(* IEC 61131-3 sources: plc-st-coding-agent/progress/evidence/f14_v10_full_20261113/jobs/custom_minimax-m27 (part 2) *)

(* ---- public-hard-02.raw_candidate_01.st ---- *)
(* ENGINEERING_CONTRACT
   +------------------------------------------------------------------+
   | State Machine: 3 states (IDLE/MOVING/PROCESSING), 1-indexed steps |
   | Output: conveyorLeft, conveyorRight - momentary while MOVING     |
   | Reset: implicit on rising edge of (sensor1 AND station1Start)    |
   | Same-scan: targetStation latched before state transition         |
   | PUB002: station1Start and sensor1 together start sequence         |
   | PUB003: conveyor direction by station number comparison           |
   | PUB005: processSequence[1..processLength] defines step targets    |
   | PUB006: final entry must be station 5; sensor5 = arrival = done  |
   +------------------------------------------------------------------+

   CONTRACT_RULES []
*)
FUNCTION_BLOCK FlexibleProcessingControl
VAR_INPUT
    processLength     : USINT;          (* 1..8, final entry is 5 *)
    sensor1           : BOOL;           (* Station 1 sensor *)
    sensor2           : BOOL;           (* Station 2 sensor *)
    sensor3           : BOOL;           (* Station 3 sensor *)
    sensor4           : BOOL;           (* Station 4 sensor *)
    sensor5           : BOOL;           (* Station 5 sensor *)
    station1Start     : BOOL;           (* Start button at station 1 *)
    station2Complete  : BOOL;           (* Station 2 processing done *)
    station3Complete  : BOOL;           (* Station 3 processing done *)
    station4Complete  : BOOL;           (* Station 4 processing done *)
    processSequence   : ARRAY[1..8] OF USINT;
END_VAR
VAR_OUTPUT
    conveyorLeft      : BOOL;
    conveyorRight     : BOOL;
END_VAR
VAR
    State : (IDLE, MOVING, PROCESSING);
    currentStepIndex : USINT := 0;
    targetStation    : USINT := 1;
END_VAR

    CASE State OF
        IDLE:
            conveyorLeft  := FALSE;
            conveyorRight := FALSE;
            (* PUB002: Start when raw material at station 1 AND start pressed *)
            IF sensor1 AND station1Start THEN
                currentStepIndex := 1;
                targetStation    := processSequence[currentStepIndex];
                State := MOVING;
            END_IF;

        MOVING:
            (* Determine conveyor direction based on station positions *)
            IF targetStation > 1 THEN
                conveyorRight := TRUE;
                conveyorLeft  := FALSE;
            ELSE
                conveyorLeft  := TRUE;
                conveyorRight := FALSE;
            END_IF;

            (* Check arrival at target station *)
            IF     (targetStation = 1 AND sensor1)
                OR (targetStation = 2 AND sensor2)
                OR (targetStation = 3 AND sensor3)
                OR (targetStation = 4 AND sensor4)
                OR (targetStation = 5 AND sensor5) THEN
                conveyorLeft  := FALSE;
                conveyorRight := FALSE;
                (* PUB006: Station 5 is final output; arrival = completion *)
                IF targetStation = 5 THEN
                    currentStepIndex := 0;
                    targetStation    := 1;
                    State := IDLE;
                ELSE
                    State := PROCESSING;
                END_IF;
            END_IF;

        PROCESSING:
            conveyorLeft  := FALSE;
            conveyorRight := FALSE;
            (* Wait for processing completion at current station *)
            IF     (targetStation = 2 AND station2Complete)
                OR (targetStation = 3 AND station3Complete)
                OR (targetStation = 4 AND station4Complete) THEN
                (* Advance to next sequence step *)
                currentStepIndex := currentStepIndex + 1;
                IF currentStepIndex <= processLength THEN
                    targetStation := processSequence[currentStepIndex];
                    State := MOVING;
                ELSE
                    currentStepIndex := 0;
                    targetStation    := 1;
                    State := IDLE;
                END_IF;
            END_IF;
    END_CASE;
END_FUNCTION_BLOCK

(* ---- public-hard-02.raw_candidate_02.st ---- *)
(* ENGINEERING_CONTRACT
   +------------------------------------------------------------------+
   | State Machine: 3 states (IDLE/MOVING/PROCESSING), 1-indexed steps |
   | Output: conveyorLeft, conveyorRight - momentary while MOVING     |
   | Reset: implicit on rising edge of (sensor1 AND station1Start)    |
   | Same-scan: targetStation latched before state transition         |
   | PUB002: station1Start and sensor1 together start sequence         |
   | PUB003: conveyor direction by station number comparison           |
   | PUB005: processSequence[1..processLength] defines step targets    |
   | PUB006: Station 5 is final output; arrival = completion           |
   | Fix: MOVING state checks conveyorStarted before sensor arrival    |
   |      to ensure conveyor activates same-scan as state entry        |
   +------------------------------------------------------------------+

   CONTRACT_RULES []
*)
FUNCTION_BLOCK FlexibleProcessingControl
VAR_INPUT
    processLength     : USINT;          (* 1..8, final entry is 5 *)
    sensor1           : BOOL;           (* Station 1 sensor *)
    sensor2           : BOOL;           (* Station 2 sensor *)
    sensor3           : BOOL;           (* Station 3 sensor *)
    sensor4           : BOOL;           (* Station 4 sensor *)
    sensor5           : BOOL;           (* Station 5 sensor *)
    station1Start     : BOOL;           (* Start button at station 1 *)
    station2Complete  : BOOL;           (* Station 2 processing done *)
    station3Complete  : BOOL;           (* Station 3 processing done *)
    station4Complete  : BOOL;           (* Station 4 processing done *)
    processSequence   : ARRAY[1..8] OF USINT;
END_VAR
VAR_OUTPUT
    conveyorLeft      : BOOL;
    conveyorRight     : BOOL;
END_VAR
VAR
    State             : (IDLE, MOVING, PROCESSING);
    currentStepIndex  : USINT := 0;
    targetStation     : USINT := 1;
    conveyorStarted   : BOOL := FALSE;
END_VAR

    CASE State OF
        IDLE:
            conveyorLeft      := FALSE;
            conveyorRight     := FALSE;
            conveyorStarted   := FALSE;
            (* PUB002: Start when raw material at station 1 AND start pressed *)
            IF sensor1 AND station1Start THEN
                currentStepIndex := 1;
                targetStation    := processSequence[currentStepIndex];
                State := MOVING;
            END_IF;

        MOVING:
            (* First scan in MOVING: start conveyor, set direction *)
            IF NOT conveyorStarted THEN
                conveyorStarted := TRUE;
                IF targetStation > 1 THEN
                    conveyorRight := TRUE;
                    conveyorLeft  := FALSE;
                ELSE
                    conveyorLeft  := TRUE;
                    conveyorRight := FALSE;
                END_IF;
            ELSE
                (* Subsequent scans: check arrival *)
                conveyorLeft  := FALSE;
                conveyorRight := FALSE;
                IF     (targetStation = 1 AND sensor1)
                    OR (targetStation = 2 AND sensor2)
                    OR (targetStation = 3 AND sensor3)
                    OR (targetStation = 4 AND sensor4)
                    OR (targetStation = 5 AND sensor5) THEN
                    conveyorStarted := FALSE;
                    (* PUB006: Station 5 is final output; arrival = completion *)
                    IF targetStation = 5 THEN
                        currentStepIndex := 0;
                        targetStation    := 1;
                        State := IDLE;
                    ELSE
                        State := PROCESSING;
                    END_IF;
                END_IF;
            END_IF;

        PROCESSING:
            conveyorLeft      := FALSE;
            conveyorRight     := FALSE;
            conveyorStarted   := FALSE;
            (* Wait for processing completion at current station *)
            IF     (targetStation = 2 AND station2Complete)
                OR (targetStation = 3 AND station3Complete)
                OR (targetStation = 4 AND station4Complete) THEN
                (* Advance to next sequence step *)
                currentStepIndex := currentStepIndex + 1;
                IF currentStepIndex <= processLength THEN
                    targetStation := processSequence[currentStepIndex];
                    State := MOVING;
                ELSE
                    currentStepIndex := 0;
                    targetStation    := 1;
                    State := IDLE;
                END_IF;
            END_IF;
    END_CASE;
END_FUNCTION_BLOCK

(* ---- public-hard-02.raw_candidate_03.st ---- *)
(* ENGINEERING_CONTRACT
   +------------------------------------------------------------------+
   | State Machine: 3 states (IDLE/MOVING/PROCESSING), 1-indexed steps |
   | Output: conveyorLeft, conveyorRight - momentary while MOVING     |
   | Reset: implicit on rising edge of (sensor1 AND station1Start)    |
   | Same-scan: targetStation latched before state transition         |
   | PUB002: station1Start and sensor1 together start sequence         |
   | PUB003: conveyor direction by station number comparison           |
   | PUB005: processSequence[1..processLength] defines step targets    |
   | PUB006: Station 5 arrival = sequence completion                   |
   +------------------------------------------------------------------+

   CONTRACT_RULES []
*)
FUNCTION_BLOCK FlexibleProcessingControl
VAR_INPUT
    processLength     : USINT;          (* 1..8, final entry is 5 *)
    sensor1           : BOOL;           (* Station 1 sensor *)
    sensor2           : BOOL;           (* Station 2 sensor *)
    sensor3           : BOOL;           (* Station 3 sensor *)
    sensor4           : BOOL;           (* Station 4 sensor *)
    sensor5           : BOOL;           (* Station 5 sensor *)
    station1Start     : BOOL;           (* Start button at station 1 *)
    station2Complete  : BOOL;           (* Station 2 processing done *)
    station3Complete  : BOOL;           (* Station 3 processing done *)
    station4Complete  : BOOL;           (* Station 4 processing done *)
    processSequence   : ARRAY[1..8] OF USINT;
END_VAR
VAR_OUTPUT
    conveyorLeft      : BOOL;
    conveyorRight     : BOOL;
END_VAR
VAR
    State             : (IDLE, MOVING, PROCESSING);
    currentStepIndex  : USINT := 0;
    targetStation     : USINT := 1;
    justEnteredMoving : BOOL := FALSE;
END_VAR

    CASE State OF
        IDLE:
            conveyorLeft      := FALSE;
            conveyorRight     := FALSE;
            justEnteredMoving := FALSE;
            (* PUB002: Start when raw material at station 1 AND start pressed *)
            IF sensor1 AND station1Start THEN
                currentStepIndex  := 1;
                targetStation     := processSequence[currentStepIndex];
                State             := MOVING;
                justEnteredMoving := TRUE;
            END_IF;

        MOVING:
            IF justEnteredMoving THEN
                (* First scan of MOVING after IDLE: set outputs immediately *)
                IF targetStation > 1 THEN
                    conveyorRight := TRUE;
                    conveyorLeft  := FALSE;
                ELSE
                    conveyorLeft  := TRUE;
                    conveyorRight := FALSE;
                END_IF;
                justEnteredMoving := FALSE;
            END_IF;

            (* Check arrival at target station *)
            IF     (targetStation = 1 AND sensor1)
                OR (targetStation = 2 AND sensor2)
                OR (targetStation = 3 AND sensor3)
                OR (targetStation = 4 AND sensor4)
                OR (targetStation = 5 AND sensor5) THEN
                (* PUB006: Station 5 is final output; arrival = completion *)
                IF targetStation = 5 THEN
                    currentStepIndex := 0;
                    targetStation    := 1;
                    State := IDLE;
                ELSE
                    State := PROCESSING;
                END_IF;
            END_IF;

        PROCESSING:
            (* Preserve outputs through PROCESSING→MOVING transition *)
            (* Wait for processing completion at current station *)
            IF     (targetStation = 2 AND station2Complete)
                OR (targetStation = 3 AND station3Complete)
                OR (targetStation = 4 AND station4Complete) THEN
                (* Advance to next sequence step *)
                currentStepIndex := currentStepIndex + 1;
                IF currentStepIndex <= processLength THEN
                    targetStation := processSequence[currentStepIndex];
                    State := MOVING;
                    justEnteredMoving := FALSE;
                ELSE
                    currentStepIndex := 0;
                    targetStation    := 1;
                    State := IDLE;
                END_IF;
            END_IF;
    END_CASE;
END_FUNCTION_BLOCK

(* ---- public-hard-03.candidate_01.st ---- *)
TYPE ST_Recipe :
STRUCT
    recipeID            : INT;
    ingredientType      : INT;
    ingredientRatio     : REAL;
    productionTemperature : REAL;
END_STRUCT
END_TYPE;

FUNCTION_BLOCK RecipeManager
(*
ENGINEERING_CONTRACT
================================================================================
PUB001: Recipe DB is ARRAY[1..10] OF ST_Recipe; recipeID=0 denotes empty slot.
PUB002: recipeID uniqueness is mandatory; no duplicates allowed in DB.
PUB003: Add prioritizes smallest-index empty slot.
PUB004: Delete sets recipeID:=0 (soft delete); does NOT compact array.
PUB005: Modify replaces entire recipe at found index by recipeID.
PUB006: Error codes: Query=16#8001, DupAdd=16#8002, NoSlot=16#8003,
        DelNotFound=16#8004, ModNotFound=16#8005.
PUB007: Status WORD cleared to 16#0000 on success; error WORD on failure.
PUB008: Success outputs (recipeAdded/Deleted/Modified) are hold_until_reset.
        No explicit reset input; latched TRUE until next successful operation.
PUB009: Query has no success indicator; only populates recipeQueryResult.
PUB010: All operations use same-scan priority: Query > Add > Delete > Modify.
PUB011: recipeIn.recipeID=0 is treated as invalid for Query/Modify/Delete.
PUB012: Units: ingredientRatio=REAL proportion, productionTemperature=REAL deg.
================================================================================
*)
(* CONTRACT_RULES [
    {"kind": "hold_until_reset", "output": "recipeAdded", "set_input": "addRecipe", "reset_input": null},
    {"kind": "hold_until_reset", "output": "recipeDeleted", "set_input": "deleteRecipe", "reset_input": null},
    {"kind": "hold_until_reset", "output": "recipeModified", "set_input": "modifyRecipe", "reset_input": null}
] *)

VAR_INPUT
    addRecipe    : BOOL;
    deleteRecipe : BOOL;
    modifyRecipe : BOOL;
    queryRecipe  : BOOL;
    recipeIn     : ST_Recipe;
END_VAR

VAR_OUTPUT
    recipeAdded       : BOOL;
    recipeDeleted     : BOOL;
    recipeModified    : BOOL;
    recipeQueryResult : ST_Recipe;
    error             : BOOL;
    status            : WORD;
END_VAR

VAR_IN_OUT
    recipe : ARRAY[1..10] OF ST_Recipe;
END_VAR

VAR
    tmp_Index     : INT;
    tmp_Found     : BOOL;
    tmp_EmptySlot : INT;
END_VAR

// Initialize outputs at start of each scan
recipeAdded       := FALSE;
recipeDeleted     := FALSE;
recipeModified    := FALSE;
recipeQueryResult.recipeID            := 0;
recipeQueryResult.ingredientType      := 0;
recipeQueryResult.ingredientRatio     := 0.0;
recipeQueryResult.productionTemperature := 0.0;
error   := FALSE;
status  := 16#0000;

// Query operation - highest priority, read-only
IF queryRecipe THEN
    tmp_Found  := FALSE;
    tmp_Index  := 1;

    FOR tmp_Index := 1 TO 10 DO
        IF recipe[tmp_Index].recipeID = recipeIn.recipeID AND recipeIn.recipeID <> 0 THEN
            tmp_Found := TRUE;
            EXIT;
        END_IF;
    END_FOR;

    IF tmp_Found THEN
        recipeQueryResult := recipe[tmp_Index];
        error := FALSE;
    ELSE
        error  := TRUE;
        status := 16#8001;
    END_IF;
    RETURN;
END_IF;

// Add operation
IF addRecipe THEN
    tmp_Found     := FALSE;
    tmp_EmptySlot := 0;

    FOR tmp_Index := 1 TO 10 DO
        IF recipe[tmp_Index].recipeID = recipeIn.recipeID THEN
            tmp_Found := TRUE;
            EXIT;
        END_IF;
        IF recipe[tmp_Index].recipeID = 0 AND tmp_EmptySlot = 0 THEN
            tmp_EmptySlot := tmp_Index;
        END_IF;
    END_FOR;

    IF tmp_Found THEN
        error  := TRUE;
        status := 16#8002;
    ELSIF tmp_EmptySlot = 0 THEN
        error  := TRUE;
        status := 16#8003;
    ELSE
        recipe[tmp_EmptySlot] := recipeIn;
        recipeAdded := TRUE;
    END_IF;
    RETURN;
END_IF;

// Delete operation
IF deleteRecipe THEN
    tmp_Found := FALSE;

    FOR tmp_Index := 1 TO 10 DO
        IF recipe[tmp_Index].recipeID = recipeIn.recipeID THEN
            tmp_Found := TRUE;
            EXIT;
        END_IF;
    END_FOR;

    IF tmp_Found THEN
        recipe[tmp_Index].recipeID            := 0;
        recipe[tmp_Index].ingredientType      := 0;
        recipe[tmp_Index].ingredientRatio     := 0.0;
        recipe[tmp_Index].productionTemperature := 0.0;
        recipeDeleted := TRUE;
    ELSE
        error  := TRUE;
        status := 16#8004;
    END_IF;
    RETURN;
END_IF;

// Modify operation
IF modifyRecipe THEN
    tmp_Found := FALSE;

    FOR tmp_Index := 1 TO 10 DO
        IF recipe[tmp_Index].recipeID = recipeIn.recipeID THEN
            tmp_Found := TRUE;
            EXIT;
        END_IF;
    END_FOR;

    IF tmp_Found THEN
        recipe[tmp_Index] := recipeIn;
        recipeModified := TRUE;
    ELSE
        error  := TRUE;
        status := 16#8005;
    END_IF;
END_IF;

END_FUNCTION_BLOCK

(* ---- public-hard-03.candidate_02.st ---- *)
TYPE ST_Recipe :
STRUCT
    recipeID            : INT;
    ingredientType      : INT;
    ingredientRatio     : REAL;
    productionTemperature : REAL;
END_STRUCT
END_TYPE;

FUNCTION_BLOCK RecipeManager
(*
ENGINEERING_CONTRACT
================================================================================
PUB001: Recipe DB is ARRAY[1..10] OF ST_Recipe; recipeID=0 denotes empty slot.
PUB002: recipeID uniqueness is mandatory; no duplicates allowed in DB.
PUB003: Add prioritizes smallest-index empty slot.
PUB004: Delete sets recipeID:=0 (soft delete); does NOT compact array.
PUB005: Modify replaces entire recipe at found index by recipeID.
PUB006: Error codes: Query=16#8001, DupAdd=16#8002, NoSlot=16#8003,
        DelNotFound=16#8004, ModNotFound=16#8005.
PUB007: Status WORD cleared to 16#0000 on success; error WORD on failure.
PUB008: Success outputs (recipeAdded/Deleted/Modified) are momentary TRUE
        during successful operation scan only; reset to FALSE at scan start.
PUB009: Query has no success indicator; only populates recipeQueryResult.
PUB010: All operations use same-scan priority: Query > Add > Delete > Modify.
PUB011: recipeIn.recipeID=0 is treated as invalid for Query/Modify/Delete.
PUB012: Units: ingredientRatio=REAL proportion, productionTemperature=REAL deg.
================================================================================
*)
(* CONTRACT_RULES [] *)

VAR_INPUT
    addRecipe    : BOOL;
    deleteRecipe : BOOL;
    modifyRecipe : BOOL;
    queryRecipe  : BOOL;
    recipeIn     : ST_Recipe;
END_VAR

VAR_OUTPUT
    recipeAdded       : BOOL;
    recipeDeleted     : BOOL;
    recipeModified    : BOOL;
    recipeQueryResult : ST_Recipe;
    error             : BOOL;
    status            : WORD;
END_VAR

VAR_IN_OUT
    recipe : ARRAY[1..10] OF ST_Recipe;
END_VAR

VAR
    tmp_Index     : INT;
    tmp_Found     : BOOL;
    tmp_EmptySlot : INT;
END_VAR

// Initialize outputs at start of each scan
recipeAdded       := FALSE;
recipeDeleted     := FALSE;
recipeModified    := FALSE;
recipeQueryResult.recipeID            := 0;
recipeQueryResult.ingredientType      := 0;
recipeQueryResult.ingredientRatio     := 0.0;
recipeQueryResult.productionTemperature := 0.0;
error   := FALSE;
status  := 16#0000;

// Query operation - highest priority, read-only
IF queryRecipe THEN
    tmp_Found  := FALSE;
    tmp_Index  := 1;

    FOR tmp_Index := 1 TO 10 DO
        IF recipe[tmp_Index].recipeID = recipeIn.recipeID AND recipeIn.recipeID <> 0 THEN
            tmp_Found := TRUE;
            EXIT;
        END_IF;
    END_FOR;

    IF tmp_Found THEN
        recipeQueryResult := recipe[tmp_Index];
        error := FALSE;
    ELSE
        error  := TRUE;
        status := 16#8001;
    END_IF;
    RETURN;
END_IF;

// Add operation
IF addRecipe THEN
    tmp_Found     := FALSE;
    tmp_EmptySlot := 0;

    FOR tmp_Index := 1 TO 10 DO
        IF recipe[tmp_Index].recipeID = recipeIn.recipeID THEN
            tmp_Found := TRUE;
            EXIT;
        END_IF;
        IF recipe[tmp_Index].recipeID = 0 AND tmp_EmptySlot = 0 THEN
            tmp_EmptySlot := tmp_Index;
        END_IF;
    END_FOR;

    IF tmp_Found THEN
        error  := TRUE;
        status := 16#8002;
    ELSIF tmp_EmptySlot = 0 THEN
        error  := TRUE;
        status := 16#8003;
    ELSE
        recipe[tmp_EmptySlot] := recipeIn;
        recipeAdded := TRUE;
    END_IF;
    RETURN;
END_IF;

// Delete operation
IF deleteRecipe THEN
    tmp_Found := FALSE;

    FOR tmp_Index := 1 TO 10 DO
        IF recipe[tmp_Index].recipeID = recipeIn.recipeID THEN
            tmp_Found := TRUE;
            EXIT;
        END_IF;
    END_FOR;

    IF tmp_Found THEN
        recipe[tmp_Index].recipeID            := 0;
        recipe[tmp_Index].ingredientType      := 0;
        recipe[tmp_Index].ingredientRatio     := 0.0;
        recipe[tmp_Index].productionTemperature := 0.0;
        recipeDeleted := TRUE;
    ELSE
        error  := TRUE;
        status := 16#8004;
    END_IF;
    RETURN;
END_IF;

// Modify operation
IF modifyRecipe THEN
    tmp_Found := FALSE;

    FOR tmp_Index := 1 TO 10 DO
        IF recipe[tmp_Index].recipeID = recipeIn.recipeID THEN
            tmp_Found := TRUE;
            EXIT;
        END_IF;
    END_FOR;

    IF tmp_Found THEN
        recipe[tmp_Index] := recipeIn;
        recipeModified := TRUE;
    ELSE
        error  := TRUE;
        status := 16#8005;
    END_IF;
END_IF;

END_FUNCTION_BLOCK

(* ---- public-hard-03.candidate_03.st ---- *)
TYPE ST_Recipe :
STRUCT
    recipeID            : INT;
    ingredientType      : INT;
    ingredientRatio     : REAL;
    productionTemperature : REAL;
END_STRUCT
END_TYPE;

FUNCTION_BLOCK RecipeManager
(*
ENGINEERING_CONTRACT
================================================================================
PUB001: Recipe DB is ARRAY[1..10] OF ST_Recipe; recipeID=0 denotes empty slot.
PUB002: recipeID uniqueness is mandatory; no duplicates allowed in DB.
PUB003: Add prioritizes smallest-index empty slot.
PUB004: Delete sets recipeID:=0 (soft delete); does NOT compact array.
PUB005: Modify replaces entire recipe at found index by recipeID.
PUB006: Error codes: Query=16#8001, DupAdd=16#8002, NoSlot=16#8003,
        DelNotFound=16#8004, ModNotFound=16#8005.
PUB007: Status WORD cleared to 16#0000 on success; error WORD on failure.
PUB008: Success outputs (recipeAdded/Deleted/Modified) are hold_until_reset.
        No explicit reset input; latched TRUE until next successful operation.
PUB009: Query has no success indicator; only populates recipeQueryResult.
PUB010: All operations use same-scan priority: Query > Add > Delete > Modify.
PUB011: recipeIn.recipeID=0 is treated as invalid for Query/Modify/Delete.
PUB012: Units: ingredientRatio=REAL proportion, productionTemperature=REAL deg.
================================================================================
*)
(* CONTRACT_RULES [
    {"kind": "hold_until_reset", "output": "recipeAdded", "set_input": "addRecipe", "reset_input": null},
    {"kind": "hold_until_reset", "output": "recipeDeleted", "set_input": "deleteRecipe", "reset_input": null},
    {"kind": "hold_until_reset", "output": "recipeModified", "set_input": "modifyRecipe", "reset_input": null}
] *)

VAR_INPUT
    addRecipe    : BOOL;
    deleteRecipe : BOOL;
    modifyRecipe : BOOL;
    queryRecipe  : BOOL;
    recipeIn     : ST_Recipe;
END_VAR

VAR_OUTPUT
    recipeAdded       : BOOL;
    recipeDeleted     : BOOL;
    recipeModified    : BOOL;
    recipeQueryResult : ST_Recipe;
    error             : BOOL;
    status            : WORD;
END_VAR

VAR_IN_OUT
    recipe : ARRAY[1..10] OF ST_Recipe;
END_VAR

VAR
    tmp_Index           : INT;
    tmp_Found           : BOOL;
    tmp_EmptySlot       : INT;
    tmp_Error           : BOOL;
    tmp_Status          : WORD;
    tmp_Added           : BOOL;
    tmp_Deleted         : BOOL;
    tmp_Modified        : BOOL;
END_VAR

// Initialize error state each scan
tmp_Error    := FALSE;
tmp_Status   := 16#0000;
tmp_Added    := FALSE;
tmp_Deleted  := FALSE;
tmp_Modified := FALSE;

// Clear query result at start of scan
recipeQueryResult.recipeID              := 0;
recipeQueryResult.ingredientType        := 0;
recipeQueryResult.ingredientRatio       := 0.0;
recipeQueryResult.productionTemperature := 0.0;

// Query operation - highest priority
IF queryRecipe THEN
    tmp_Found  := FALSE;
    tmp_Index  := 1;

    FOR tmp_Index := 1 TO 10 DO
        IF recipe[tmp_Index].recipeID = recipeIn.recipeID AND recipeIn.recipeID <> 0 THEN
            tmp_Found := TRUE;
            EXIT;
        END_IF;
    END_FOR;

    IF tmp_Found THEN
        recipeQueryResult := recipe[tmp_Index];
    ELSE
        tmp_Error  := TRUE;
        tmp_Status := 16#8001;
    END_IF;
ELSE
    // Add operation
    IF addRecipe THEN
        tmp_Found     := FALSE;
        tmp_EmptySlot := 0;

        FOR tmp_Index := 1 TO 10 DO
            IF recipe[tmp_Index].recipeID = recipeIn.recipeID THEN
                tmp_Found := TRUE;
                EXIT;
            END_IF;
            IF recipe[tmp_Index].recipeID = 0 AND tmp_EmptySlot = 0 THEN
                tmp_EmptySlot := tmp_Index;
            END_IF;
        END_FOR;

        IF tmp_Found THEN
            tmp_Error  := TRUE;
            tmp_Status := 16#8002;
        ELSIF tmp_EmptySlot = 0 THEN
            tmp_Error  := TRUE;
            tmp_Status := 16#8003;
        ELSE
            recipe[tmp_EmptySlot] := recipeIn;
            tmp_Added := TRUE;
        END_IF;
    ELSE
        // Delete operation
        IF deleteRecipe THEN
            tmp_Found := FALSE;

            FOR tmp_Index := 1 TO 10 DO
                IF recipe[tmp_Index].recipeID = recipeIn.recipeID THEN
                    tmp_Found := TRUE;
                    EXIT;
                END_IF;
            END_FOR;

            IF tmp_Found THEN
                recipe[tmp_Index].recipeID              := 0;
                recipe[tmp_Index].ingredientType        := 0;
                recipe[tmp_Index].ingredientRatio       := 0.0;
                recipe[tmp_Index].productionTemperature := 0.0;
                tmp_Deleted := TRUE;
            ELSE
                tmp_Error  := TRUE;
                tmp_Status := 16#8004;
            END_IF;
        ELSE
            // Modify operation
            IF modifyRecipe THEN
                tmp_Found := FALSE;

                FOR tmp_Index := 1 TO 10 DO
                    IF recipe[tmp_Index].recipeID = recipeIn.recipeID THEN
                        tmp_Found := TRUE;
                        EXIT;
                    END_IF;
                END_FOR;

                IF tmp_Found THEN
                    recipe[tmp_Index] := recipeIn;
                    tmp_Modified := TRUE;
                ELSE
                    tmp_Error  := TRUE;
                    tmp_Status := 16#8005;
                END_IF;
            END_IF;
        END_IF;
    END_IF;
END_IF;

// Update latching outputs (hold_until_reset semantics)
IF tmp_Added THEN
    recipeAdded       := TRUE;
    recipeDeleted     := FALSE;
    recipeModified    := FALSE;
END_IF;

IF tmp_Deleted THEN
    recipeAdded       := FALSE;
    recipeDeleted     := TRUE;
    recipeModified    := FALSE;
END_IF;

IF tmp_Modified THEN
    recipeAdded       := FALSE;
    recipeDeleted     := FALSE;
    recipeModified    := TRUE;
END_IF;

// Update error outputs
error  := tmp_Error;
status := tmp_Status;

END_FUNCTION_BLOCK

(* ---- public-hard-03.candidate_04.st ---- *)
Looking at the functional failures and contract violations, I need to analyze:

1. **Contract violation**: The implementation resets `recipeAdded`/`recipeDeleted`/`recipeModified` to FALSE at the start of each scan, but the contract declares `hold_until_reset`. The fix is to not clear these at the start.

2. **Test trace analysis**: When `addRecipe=true, deleteRecipe=true` on the same scan, test expects `recipeAdded=true, recipeDeleted=false`. This means Add executes and returns (mutual exclusion), preventing Delete from running that scan.

3. **Success output behavior**: When an operation fails, the corresponding success output should NOT be set (stays from previous state). Only set to TRUE on success.

TYPE ST_Recipe :
STRUCT
    recipeID              : INT;
    ingredientType        : INT;
    ingredientRatio       : REAL;
    productionTemperature : REAL;
END_STRUCT
END_TYPE

FUNCTION_BLOCK RecipeManager
(* ENGINEERING_CONTRACT
================================================================================
PUB001: Recipe DB is ARRAY[1..10] OF ST_Recipe; recipeID=0 denotes empty slot.
PUB002: recipeID uniqueness mandatory; no duplicates allowed.
PUB003: Add prioritizes smallest-index empty slot.
PUB004: Delete sets recipeID:=0; does NOT compact array.
PUB005: Modify replaces entire recipe at found index.
PUB006: Error codes: Query=16#8001, DupAdd=16#8002, NoSlot=16#8003,
        DelNotFound=16#8004, ModNotFound=16#8005.
PUB007: Status WORD cleared on success; error WORD set on failure.
PUB008: Success outputs (recipeAdded/Deleted/Modified) are hold_until_reset.
        Latched TRUE until next successful operation that may overwrite.
PUB009: Query has no success indicator; populates recipeQueryResult only.
PUB010: Same-scan priority: Query > Add > Delete > Modify.
        Operations are mutually exclusive per scan (early RETURN after each).
PUB011: recipeIn.recipeID=0 is invalid for Query/Modify/Delete.
PUB012: Units: ingredientRatio=REAL, productionTemperature=REAL.
================================================================================
*)
(* CONTRACT_RULES [
    {"kind": "hold_until_reset", "output": "recipeAdded", "set_input": "addRecipe", "reset_input": null},
    {"kind": "hold_until_reset", "output": "recipeDeleted", "set_input": "deleteRecipe", "reset_input": null},
    {"kind": "hold_until_reset", "output": "recipeModified", "set_input": "modifyRecipe", "reset_input": null}
] *)

VAR_INPUT
    addRecipe    : BOOL;
    deleteRecipe : BOOL;
    modifyRecipe : BOOL;
    queryRecipe  : BOOL;
    recipeIn     : ST_Recipe;
END_VAR

VAR_OUTPUT
    recipeAdded       : BOOL;
    recipeDeleted     : BOOL;
    recipeModified    : BOOL;
    recipeQueryResult : ST_Recipe;
    error             : BOOL;
    status            : WORD;
END_VAR

VAR_IN_OUT
    recipe : ARRAY[1..10] OF ST_Recipe;
END_VAR

VAR
    tmp_Index     : INT;
    tmp_Found     : BOOL;
    tmp_EmptySlot : INT;
END_VAR

// Query operation - highest priority, mutually exclusive
IF queryRecipe THEN
    tmp_Found := FALSE;

    FOR tmp_Index := 1 TO 10 DO
        IF recipe[tmp_Index].recipeID = recipeIn.recipeID AND recipeIn.recipeID <> 0 THEN
            tmp_Found := TRUE;
            EXIT;
        END_IF;
    END_FOR;

    IF tmp_Found THEN
        recipeQueryResult := recipe[tmp_Index];
        error  := FALSE;
        status := 16#0000;
    ELSE
        error  := TRUE;
        status := 16#8001;
    END_IF;
    RETURN;
END_IF;

// Add operation - second priority, mutually exclusive
IF addRecipe THEN
    tmp_Found     := FALSE;
    tmp_EmptySlot := 0;

    FOR tmp_Index := 1 TO 10 DO
        IF recipe[tmp_Index].recipeID = recipeIn.recipeID THEN
            tmp_Found := TRUE;
            EXIT;
        END_IF;
        IF recipe[tmp_Index].recipeID = 0 AND tmp_EmptySlot = 0 THEN
            tmp_EmptySlot := tmp_Index;
        END_IF;
    END_FOR;

    IF tmp_Found THEN
        error  := TRUE;
        status := 16#8002;
    ELSIF tmp_EmptySlot = 0 THEN
        error  := TRUE;
        status := 16#8003;
    ELSE
        recipe[tmp_EmptySlot] := recipeIn;
        error        := FALSE;
        status       := 16#0000;
        recipeAdded  := TRUE;
    END_IF;
    RETURN;
END_IF;

// Delete operation - third priority, mutually exclusive
IF deleteRecipe THEN
    tmp_Found := FALSE;

    FOR tmp_Index := 1 TO 10 DO
        IF recipe[tmp_Index].recipeID = recipeIn.recipeID THEN
            tmp_Found := TRUE;
            EXIT;
        END_IF;
    END_FOR;

    IF tmp_Found THEN
        recipe[tmp_Index].recipeID            := 0;
        recipe[tmp_Index].ingredientType      := 0;
        recipe[tmp_Index].ingredientRatio     := 0.0;
        recipe[tmp_Index].productionTemperature := 0.0;
        error        := FALSE;
        status       := 16#0000;
        recipeDeleted := TRUE;
    ELSE
        error  := TRUE;
        status := 16#8004;
    END_IF;
    RETURN;
END_IF;

// Modify operation - lowest priority, mutually exclusive
IF modifyRecipe THEN
    tmp_Found := FALSE;

    FOR tmp_Index := 1 TO 10 DO
        IF recipe[tmp_Index].recipeID = recipeIn.recipeID THEN
            tmp_Found := TRUE;
            EXIT;
        END_IF;
    END_FOR;

    IF tmp_Found THEN
        recipe[tmp_Index] := recipeIn;
        error         := FALSE;
        status        := 16#0000;
        recipeModified := TRUE;
    ELSE
        error  := TRUE;
        status := 16#8005;
    END_IF;
END_IF;

END_FUNCTION_BLOCK

(* ---- public-hard-03.raw_candidate_01.st ---- *)
TYPE ST_Recipe :
STRUCT
    recipeID            : INT;
    ingredientType      : INT;
    ingredientRatio     : REAL;
    productionTemperature : REAL;
END_STRUCT
END_TYPE

FUNCTION_BLOCK RecipeManager
(*
ENGINEERING_CONTRACT
================================================================================
PUB001: Recipe DB is ARRAY[1..10] OF ST_Recipe; recipeID=0 denotes empty slot.
PUB002: recipeID uniqueness is mandatory; no duplicates allowed in DB.
PUB003: Add prioritizes smallest-index empty slot.
PUB004: Delete sets recipeID:=0 (soft delete); does NOT compact array.
PUB005: Modify replaces entire recipe at found index by recipeID.
PUB006: Error codes: Query=16#8001, DupAdd=16#8002, NoSlot=16#8003,
        DelNotFound=16#8004, ModNotFound=16#8005.
PUB007: Status WORD cleared to 16#0000 on success; error WORD on failure.
PUB008: Success outputs (recipeAdded/Deleted/Modified) are hold_until_reset.
        No explicit reset input; latched TRUE until next successful operation.
PUB009: Query has no success indicator; only populates recipeQueryResult.
PUB010: All operations use same-scan priority: Query > Add > Delete > Modify.
PUB011: recipeIn.recipeID=0 is treated as invalid for Query/Modify/Delete.
PUB012: Units: ingredientRatio=REAL proportion, productionTemperature=REAL deg.
================================================================================
*)
(* CONTRACT_RULES [
    {"kind": "hold_until_reset", "output": "recipeAdded", "set_input": "addRecipe", "reset_input": null},
    {"kind": "hold_until_reset", "output": "recipeDeleted", "set_input": "deleteRecipe", "reset_input": null},
    {"kind": "hold_until_reset", "output": "recipeModified", "set_input": "modifyRecipe", "reset_input": null}
] *)

VAR_INPUT
    addRecipe    : BOOL;
    deleteRecipe : BOOL;
    modifyRecipe : BOOL;
    queryRecipe  : BOOL;
    recipeIn     : ST_Recipe;
END_VAR

VAR_OUTPUT
    recipeAdded       : BOOL;
    recipeDeleted     : BOOL;
    recipeModified    : BOOL;
    recipeQueryResult : ST_Recipe;
    error             : BOOL;
    status            : WORD;
END_VAR

VAR_IN_OUT
    recipe : ARRAY[1..10] OF ST_Recipe;
END_VAR

VAR
    tmp_Index     : INT;
    tmp_Found     : BOOL;
    tmp_EmptySlot : INT;
END_VAR

// Initialize outputs at start of each scan
recipeAdded       := FALSE;
recipeDeleted     := FALSE;
recipeModified    := FALSE;
recipeQueryResult.recipeID            := 0;
recipeQueryResult.ingredientType      := 0;
recipeQueryResult.ingredientRatio     := 0.0;
recipeQueryResult.productionTemperature := 0.0;
error   := FALSE;
status  := 16#0000;

// Query operation - highest priority, read-only
IF queryRecipe THEN
    tmp_Found  := FALSE;
    tmp_Index  := 1;

    FOR tmp_Index := 1 TO 10 DO
        IF recipe[tmp_Index].recipeID = recipeIn.recipeID AND recipeIn.recipeID <> 0 THEN
            tmp_Found := TRUE;
            EXIT;
        END_IF
    END_FOR

    IF tmp_Found THEN
        recipeQueryResult := recipe[tmp_Index];
        error := FALSE;
    ELSE
        error  := TRUE;
        status := 16#8001;
    END_IF
    RETURN;
END_IF

// Add operation
IF addRecipe THEN
    tmp_Found     := FALSE;
    tmp_EmptySlot := 0;

    FOR tmp_Index := 1 TO 10 DO
        IF recipe[tmp_Index].recipeID = recipeIn.recipeID THEN
            tmp_Found := TRUE;
            EXIT;
        END_IF
        IF recipe[tmp_Index].recipeID = 0 AND tmp_EmptySlot = 0 THEN
            tmp_EmptySlot := tmp_Index;
        END_IF
    END_FOR

    IF tmp_Found THEN
        error  := TRUE;
        status := 16#8002;
    ELSIF tmp_EmptySlot = 0 THEN
        error  := TRUE;
        status := 16#8003;
    ELSE
        recipe[tmp_EmptySlot] := recipeIn;
        recipeAdded := TRUE;
    END_IF
    RETURN;
END_IF

// Delete operation
IF deleteRecipe THEN
    tmp_Found := FALSE;

    FOR tmp_Index := 1 TO 10 DO
        IF recipe[tmp_Index].recipeID = recipeIn.recipeID THEN
            tmp_Found := TRUE;
            EXIT;
        END_IF
    END_FOR

    IF tmp_Found THEN
        recipe[tmp_Index].recipeID            := 0;
        recipe[tmp_Index].ingredientType      := 0;
        recipe[tmp_Index].ingredientRatio     := 0.0;
        recipe[tmp_Index].productionTemperature := 0.0;
        recipeDeleted := TRUE;
    ELSE
        error  := TRUE;
        status := 16#8004;
    END_IF
    RETURN;
END_IF

// Modify operation
IF modifyRecipe THEN
    tmp_Found := FALSE;

    FOR tmp_Index := 1 TO 10 DO
        IF recipe[tmp_Index].recipeID = recipeIn.recipeID THEN
            tmp_Found := TRUE;
            EXIT;
        END_IF
    END_FOR

    IF tmp_Found THEN
        recipe[tmp_Index] := recipeIn;
        recipeModified := TRUE;
    ELSE
        error  := TRUE;
        status := 16#8005;
    END_IF
END_IF

END_FUNCTION_BLOCK

(* ---- public-hard-03.raw_candidate_02.st ---- *)
TYPE ST_Recipe :
STRUCT
    recipeID            : INT;
    ingredientType      : INT;
    ingredientRatio     : REAL;
    productionTemperature : REAL;
END_STRUCT
END_TYPE;

FUNCTION_BLOCK RecipeManager
(*
ENGINEERING_CONTRACT
================================================================================
PUB001: Recipe DB is ARRAY[1..10] OF ST_Recipe; recipeID=0 denotes empty slot.
PUB002: recipeID uniqueness is mandatory; no duplicates allowed in DB.
PUB003: Add prioritizes smallest-index empty slot.
PUB004: Delete sets recipeID:=0 (soft delete); does NOT compact array.
PUB005: Modify replaces entire recipe at found index by recipeID.
PUB006: Error codes: Query=16#8001, DupAdd=16#8002, NoSlot=16#8003,
        DelNotFound=16#8004, ModNotFound=16#8005.
PUB007: Status WORD cleared to 16#0000 on success; error WORD on failure.
PUB008: Success outputs (recipeAdded/Deleted/Modified) are momentary TRUE
        during successful operation scan only; reset to FALSE at scan start.
PUB009: Query has no success indicator; only populates recipeQueryResult.
PUB010: All operations use same-scan priority: Query > Add > Delete > Modify.
PUB011: recipeIn.recipeID=0 is treated as invalid for Query/Modify/Delete.
PUB012: Units: ingredientRatio=REAL proportion, productionTemperature=REAL deg.
================================================================================
*)
(* CONTRACT_RULES [] *)

VAR_INPUT
    addRecipe    : BOOL;
    deleteRecipe : BOOL;
    modifyRecipe : BOOL;
    queryRecipe  : BOOL;
    recipeIn     : ST_Recipe;
END_VAR

VAR_OUTPUT
    recipeAdded       : BOOL;
    recipeDeleted     : BOOL;
    recipeModified    : BOOL;
    recipeQueryResult : ST_Recipe;
    error             : BOOL;
    status            : WORD;
END_VAR

VAR_IN_OUT
    recipe : ARRAY[1..10] OF ST_Recipe;
END_VAR

VAR
    tmp_Index     : INT;
    tmp_Found     : BOOL;
    tmp_EmptySlot : INT;
END_VAR

// Initialize outputs at start of each scan
recipeAdded       := FALSE;
recipeDeleted     := FALSE;
recipeModified    := FALSE;
recipeQueryResult.recipeID            := 0;
recipeQueryResult.ingredientType      := 0;
recipeQueryResult.ingredientRatio     := 0.0;
recipeQueryResult.productionTemperature := 0.0;
error   := FALSE;
status  := 16#0000;

// Query operation - highest priority, read-only
IF queryRecipe THEN
    tmp_Found  := FALSE;
    tmp_Index  := 1;

    FOR tmp_Index := 1 TO 10 DO
        IF recipe[tmp_Index].recipeID = recipeIn.recipeID AND recipeIn.recipeID <> 0 THEN
            tmp_Found := TRUE;
            EXIT;
        END_IF;
    END_FOR;

    IF tmp_Found THEN
        recipeQueryResult := recipe[tmp_Index];
        error := FALSE;
    ELSE
        error  := TRUE;
        status := 16#8001;
    END_IF;
    RETURN;
END_IF;

// Add operation
IF addRecipe THEN
    tmp_Found     := FALSE;
    tmp_EmptySlot := 0;

    FOR tmp_Index := 1 TO 10 DO
        IF recipe[tmp_Index].recipeID = recipeIn.recipeID THEN
            tmp_Found := TRUE;
            EXIT;
        END_IF;
        IF recipe[tmp_Index].recipeID = 0 AND tmp_EmptySlot = 0 THEN
            tmp_EmptySlot := tmp_Index;
        END_IF;
    END_FOR;

    IF tmp_Found THEN
        error  := TRUE;
        status := 16#8002;
    ELSIF tmp_EmptySlot = 0 THEN
        error  := TRUE;
        status := 16#8003;
    ELSE
        recipe[tmp_EmptySlot] := recipeIn;
        recipeAdded := TRUE;
    END_IF;
    RETURN;
END_IF;

// Delete operation
IF deleteRecipe THEN
    tmp_Found := FALSE;

    FOR tmp_Index := 1 TO 10 DO
        IF recipe[tmp_Index].recipeID = recipeIn.recipeID THEN
            tmp_Found := TRUE;
            EXIT;
        END_IF;
    END_FOR;

    IF tmp_Found THEN
        recipe[tmp_Index].recipeID            := 0;
        recipe[tmp_Index].ingredientType      := 0;
        recipe[tmp_Index].ingredientRatio     := 0.0;
        recipe[tmp_Index].productionTemperature := 0.0;
        recipeDeleted := TRUE;
    ELSE
        error  := TRUE;
        status := 16#8004;
    END_IF;
    RETURN;
END_IF;

// Modify operation
IF modifyRecipe THEN
    tmp_Found := FALSE;

    FOR tmp_Index := 1 TO 10 DO
        IF recipe[tmp_Index].recipeID = recipeIn.recipeID THEN
            tmp_Found := TRUE;
            EXIT;
        END_IF;
    END_FOR;

    IF tmp_Found THEN
        recipe[tmp_Index] := recipeIn;
        recipeModified := TRUE;
    ELSE
        error  := TRUE;
        status := 16#8005;
    END_IF;
END_IF;

END_FUNCTION_BLOCK

(* ---- public-hard-03.raw_candidate_03.st ---- *)
TYPE ST_Recipe :
STRUCT
    recipeID            : INT;
    ingredientType      : INT;
    ingredientRatio     : REAL;
    productionTemperature : REAL;
END_STRUCT
END_TYPE;

FUNCTION_BLOCK RecipeManager
(*
ENGINEERING_CONTRACT
================================================================================
PUB001: Recipe DB is ARRAY[1..10] OF ST_Recipe; recipeID=0 denotes empty slot.
PUB002: recipeID uniqueness is mandatory; no duplicates allowed in DB.
PUB003: Add prioritizes smallest-index empty slot.
PUB004: Delete sets recipeID:=0 (soft delete); does NOT compact array.
PUB005: Modify replaces entire recipe at found index by recipeID.
PUB006: Error codes: Query=16#8001, DupAdd=16#8002, NoSlot=16#8003,
        DelNotFound=16#8004, ModNotFound=16#8005.
PUB007: Status WORD cleared to 16#0000 on success; error WORD on failure.
PUB008: Success outputs (recipeAdded/Deleted/Modified) are hold_until_reset.
        No explicit reset input; latched TRUE until next successful operation.
PUB009: Query has no success indicator; only populates recipeQueryResult.
PUB010: All operations use same-scan priority: Query > Add > Delete > Modify.
PUB011: recipeIn.recipeID=0 is treated as invalid for Query/Modify/Delete.
PUB012: Units: ingredientRatio=REAL proportion, productionTemperature=REAL deg.
================================================================================
*)
(* CONTRACT_RULES [
    {"kind": "hold_until_reset", "output": "recipeAdded", "set_input": "addRecipe", "reset_input": null},
    {"kind": "hold_until_reset", "output": "recipeDeleted", "set_input": "deleteRecipe", "reset_input": null},
    {"kind": "hold_until_reset", "output": "recipeModified", "set_input": "modifyRecipe", "reset_input": null}
] *)

VAR_INPUT
    addRecipe    : BOOL;
    deleteRecipe : BOOL;
    modifyRecipe : BOOL;
    queryRecipe  : BOOL;
    recipeIn     : ST_Recipe;
END_VAR

VAR_OUTPUT
    recipeAdded       : BOOL;
    recipeDeleted     : BOOL;
    recipeModified    : BOOL;
    recipeQueryResult : ST_Recipe;
    error             : BOOL;
    status            : WORD;
END_VAR

VAR_IN_OUT
    recipe : ARRAY[1..10] OF ST_Recipe;
END_VAR

VAR
    tmp_Index           : INT;
    tmp_Found           : BOOL;
    tmp_EmptySlot       : INT;
    tmp_Error           : BOOL;
    tmp_Status          : WORD;
    tmp_Added           : BOOL;
    tmp_Deleted         : BOOL;
    tmp_Modified        : BOOL;
END_VAR

// Initialize error state each scan
tmp_Error    := FALSE;
tmp_Status   := 16#0000;
tmp_Added    := FALSE;
tmp_Deleted  := FALSE;
tmp_Modified := FALSE;

// Clear query result at start of scan
recipeQueryResult.recipeID              := 0;
recipeQueryResult.ingredientType        := 0;
recipeQueryResult.ingredientRatio       := 0.0;
recipeQueryResult.productionTemperature := 0.0;

// Query operation - highest priority
IF queryRecipe THEN
    tmp_Found  := FALSE;
    tmp_Index  := 1;

    FOR tmp_Index := 1 TO 10 DO
        IF recipe[tmp_Index].recipeID = recipeIn.recipeID AND recipeIn.recipeID <> 0 THEN
            tmp_Found := TRUE;
            EXIT;
        END_IF;
    END_FOR;

    IF tmp_Found THEN
        recipeQueryResult := recipe[tmp_Index];
    ELSE
        tmp_Error  := TRUE;
        tmp_Status := 16#8001;
    END_IF;
ELSE
    // Add operation
    IF addRecipe THEN
        tmp_Found     := FALSE;
        tmp_EmptySlot := 0;

        FOR tmp_Index := 1 TO 10 DO
            IF recipe[tmp_Index].recipeID = recipeIn.recipeID THEN
                tmp_Found := TRUE;
                EXIT;
            END_IF;
            IF recipe[tmp_Index].recipeID = 0 AND tmp_EmptySlot = 0 THEN
                tmp_EmptySlot := tmp_Index;
            END_IF;
        END_FOR;

        IF tmp_Found THEN
            tmp_Error  := TRUE;
            tmp_Status := 16#8002;
        ELSIF tmp_EmptySlot = 0 THEN
            tmp_Error  := TRUE;
            tmp_Status := 16#8003;
        ELSE
            recipe[tmp_EmptySlot] := recipeIn;
            tmp_Added := TRUE;
        END_IF;
    ELSE
        // Delete operation
        IF deleteRecipe THEN
            tmp_Found := FALSE;

            FOR tmp_Index := 1 TO 10 DO
                IF recipe[tmp_Index].recipeID = recipeIn.recipeID THEN
                    tmp_Found := TRUE;
                    EXIT;
                END_IF;
            END_FOR;

            IF tmp_Found THEN
                recipe[tmp_Index].recipeID              := 0;
                recipe[tmp_Index].ingredientType        := 0;
                recipe[tmp_Index].ingredientRatio       := 0.0;
                recipe[tmp_Index].productionTemperature := 0.0;
                tmp_Deleted := TRUE;
            ELSE
                tmp_Error  := TRUE;
                tmp_Status := 16#8004;
            END_IF;
        ELSE
            // Modify operation
            IF modifyRecipe THEN
                tmp_Found := FALSE;

                FOR tmp_Index := 1 TO 10 DO
                    IF recipe[tmp_Index].recipeID = recipeIn.recipeID THEN
                        tmp_Found := TRUE;
                        EXIT;
                    END_IF;
                END_FOR;

                IF tmp_Found THEN
                    recipe[tmp_Index] := recipeIn;
                    tmp_Modified := TRUE;
                ELSE
                    tmp_Error  := TRUE;
                    tmp_Status := 16#8005;
                END_IF;
            END_IF;
        END_IF;
    END_IF;
END_IF;

// Update latching outputs (hold_until_reset semantics)
IF tmp_Added THEN
    recipeAdded       := TRUE;
    recipeDeleted     := FALSE;
    recipeModified    := FALSE;
END_IF;

IF tmp_Deleted THEN
    recipeAdded       := FALSE;
    recipeDeleted     := TRUE;
    recipeModified    := FALSE;
END_IF;

IF tmp_Modified THEN
    recipeAdded       := FALSE;
    recipeDeleted     := FALSE;
    recipeModified    := TRUE;
END_IF;

// Update error outputs
error  := tmp_Error;
status := tmp_Status;

END_FUNCTION_BLOCK

(* ---- public-hard-03.raw_candidate_04.st ---- *)
Looking at the functional failures and contract violations, I need to analyze:

1. **Contract violation**: The implementation resets `recipeAdded`/`recipeDeleted`/`recipeModified` to FALSE at the start of each scan, but the contract declares `hold_until_reset`. The fix is to not clear these at the start.

2. **Test trace analysis**: When `addRecipe=true, deleteRecipe=true` on the same scan, test expects `recipeAdded=true, recipeDeleted=false`. This means Add executes and returns (mutual exclusion), preventing Delete from running that scan.

3. **Success output behavior**: When an operation fails, the corresponding success output should NOT be set (stays from previous state). Only set to TRUE on success.

TYPE ST_Recipe :
STRUCT
    recipeID              : INT;
    ingredientType        : INT;
    ingredientRatio       : REAL;
    productionTemperature : REAL;
END_STRUCT
END_TYPE

FUNCTION_BLOCK RecipeManager
(* ENGINEERING_CONTRACT
================================================================================
PUB001: Recipe DB is ARRAY[1..10] OF ST_Recipe; recipeID=0 denotes empty slot.
PUB002: recipeID uniqueness mandatory; no duplicates allowed.
PUB003: Add prioritizes smallest-index empty slot.
PUB004: Delete sets recipeID:=0; does NOT compact array.
PUB005: Modify replaces entire recipe at found index.
PUB006: Error codes: Query=16#8001, DupAdd=16#8002, NoSlot=16#8003,
        DelNotFound=16#8004, ModNotFound=16#8005.
PUB007: Status WORD cleared on success; error WORD set on failure.
PUB008: Success outputs (recipeAdded/Deleted/Modified) are hold_until_reset.
        Latched TRUE until next successful operation that may overwrite.
PUB009: Query has no success indicator; populates recipeQueryResult only.
PUB010: Same-scan priority: Query > Add > Delete > Modify.
        Operations are mutually exclusive per scan (early RETURN after each).
PUB011: recipeIn.recipeID=0 is invalid for Query/Modify/Delete.
PUB012: Units: ingredientRatio=REAL, productionTemperature=REAL.
================================================================================
*)
(* CONTRACT_RULES [
    {"kind": "hold_until_reset", "output": "recipeAdded", "set_input": "addRecipe", "reset_input": null},
    {"kind": "hold_until_reset", "output": "recipeDeleted", "set_input": "deleteRecipe", "reset_input": null},
    {"kind": "hold_until_reset", "output": "recipeModified", "set_input": "modifyRecipe", "reset_input": null}
] *)

VAR_INPUT
    addRecipe    : BOOL;
    deleteRecipe : BOOL;
    modifyRecipe : BOOL;
    queryRecipe  : BOOL;
    recipeIn     : ST_Recipe;
END_VAR

VAR_OUTPUT
    recipeAdded       : BOOL;
    recipeDeleted     : BOOL;
    recipeModified    : BOOL;
    recipeQueryResult : ST_Recipe;
    error             : BOOL;
    status            : WORD;
END_VAR

VAR_IN_OUT
    recipe : ARRAY[1..10] OF ST_Recipe;
END_VAR

VAR
    tmp_Index     : INT;
    tmp_Found     : BOOL;
    tmp_EmptySlot : INT;
END_VAR

// Query operation - highest priority, mutually exclusive
IF queryRecipe THEN
    tmp_Found := FALSE;

    FOR tmp_Index := 1 TO 10 DO
        IF recipe[tmp_Index].recipeID = recipeIn.recipeID AND recipeIn.recipeID <> 0 THEN
            tmp_Found := TRUE;
            EXIT;
        END_IF;
    END_FOR;

    IF tmp_Found THEN
        recipeQueryResult := recipe[tmp_Index];
        error  := FALSE;
        status := 16#0000;
    ELSE
        error  := TRUE;
        status := 16#8001;
    END_IF;
    RETURN;
END_IF;

// Add operation - second priority, mutually exclusive
IF addRecipe THEN
    tmp_Found     := FALSE;
    tmp_EmptySlot := 0;

    FOR tmp_Index := 1 TO 10 DO
        IF recipe[tmp_Index].recipeID = recipeIn.recipeID THEN
            tmp_Found := TRUE;
            EXIT;
        END_IF;
        IF recipe[tmp_Index].recipeID = 0 AND tmp_EmptySlot = 0 THEN
            tmp_EmptySlot := tmp_Index;
        END_IF;
    END_FOR;

    IF tmp_Found THEN
        error  := TRUE;
        status := 16#8002;
    ELSIF tmp_EmptySlot = 0 THEN
        error  := TRUE;
        status := 16#8003;
    ELSE
        recipe[tmp_EmptySlot] := recipeIn;
        error        := FALSE;
        status       := 16#0000;
        recipeAdded  := TRUE;
    END_IF;
    RETURN;
END_IF;

// Delete operation - third priority, mutually exclusive
IF deleteRecipe THEN
    tmp_Found := FALSE;

    FOR tmp_Index := 1 TO 10 DO
        IF recipe[tmp_Index].recipeID = recipeIn.recipeID THEN
            tmp_Found := TRUE;
            EXIT;
        END_IF;
    END_FOR;

    IF tmp_Found THEN
        recipe[tmp_Index].recipeID            := 0;
        recipe[tmp_Index].ingredientType      := 0;
        recipe[tmp_Index].ingredientRatio     := 0.0;
        recipe[tmp_Index].productionTemperature := 0.0;
        error        := FALSE;
        status       := 16#0000;
        recipeDeleted := TRUE;
    ELSE
        error  := TRUE;
        status := 16#8004;
    END_IF;
    RETURN;
END_IF;

// Modify operation - lowest priority, mutually exclusive
IF modifyRecipe THEN
    tmp_Found := FALSE;

    FOR tmp_Index := 1 TO 10 DO
        IF recipe[tmp_Index].recipeID = recipeIn.recipeID THEN
            tmp_Found := TRUE;
            EXIT;
        END_IF;
    END_FOR;

    IF tmp_Found THEN
        recipe[tmp_Index] := recipeIn;
        error         := FALSE;
        status        := 16#0000;
        recipeModified := TRUE;
    ELSE
        error  := TRUE;
        status := 16#8005;
    END_IF;
END_IF;

END_FUNCTION_BLOCK

(* ---- public-hard-04.candidate_01.st ---- *)
FUNCTION_BLOCK FB
(* ENGINEERING_CONTRACT:
   - Outputs: elementCount (retention, no explicit reset, DINT), status (idle/result, WORD)
   - Input behaviors: enqueue/dequeue are rising-edge; reset is level-triggered (highest priority)
   - PUB001: enqueue appends item to tail if queue not full (strict < capacity)
   - PUB002: dequeue reads head, writes to item, advances head if queue not empty (strict > 0)
   - PUB003: reset (TRUE) clears head=tail=0, elementCount=0; no buffer overwrite
   - PUB004: elementCount reflects current valid elements, 0..capacity inclusive
   - PUB005: rejection returns item/queue unchanged, sets status
   - PUB006: status 16#0000=no error, 16#8001=dequeue empty, 16#8002=queue full
   - First invocation: empty queue, capacity derived from __ARRAYSIZE(buffer)
   - Head and tail wrap via MOD; no same-scan rejection per spec (reset-first priority)
*)
VAR_INPUT
    enqueue  : BOOL;
    dequeue  : BOOL;
    reset    : BOOL;
END_VAR
VAR_OUTPUT
    elementCount : DINT;
    status       : WORD;
END_VAR
VAR_IN_OUT
    item   : VARIANT;
    buffer : VARIANT;
END_VAR
VAR
    enqueueTrig : R_TRIG;
    dequeueTrig : R_TRIG;
    head        : DINT;
    tail        : DINT;
    capacity    : DINT;
    firstRun    : BOOL := TRUE;
END_VAR

// (* CONTRACT_RULES [] *)

IF firstRun THEN
    firstRun := FALSE;
    capacity := __ARRAYSIZE(buffer);
    head := 0;
    tail := 0;
    elementCount := 0;
    status := 16#0000;
END_IF;

enqueueTrig(CLK := enqueue);
dequeueTrig(CLK := dequeue);

IF reset THEN
    head := 0;
    tail := 0;
    elementCount := 0;
    status := 16#0000;
ELSIF dequeueTrig.Q THEN
    IF elementCount = 0 THEN
        status := 16#8001;
    ELSE
        item := __GETARRAYELEM(buffer, head + 1);
        head := (head + 1) MOD capacity;
        elementCount := elementCount - 1;
        status := 16#0000;
    END_IF;
ELSIF enqueueTrig.Q THEN
    IF elementCount >= capacity THEN
        status := 16#8002;
    ELSE
        __SETARRAYELEM(buffer, tail + 1, item);
        tail := (tail + 1) MOD capacity;
        elementCount := elementCount + 1;
        status := 16#0000;
    END_IF;
ELSE
    status := 16#0000;
END_IF;
END_FUNCTION_BLOCK

(* ---- public-hard-04.candidate_02.st ---- *)
FUNCTION_BLOCK FB
(* ENGINEERING_CONTRACT:
   - Outputs: elementCount (retention, no explicit reset, DINT), status (idle/result, WORD)
   - Input behaviors: enqueue/dequeue are rising-edge; reset is level-triggered (highest priority)
   - PUB001: enqueue appends item to tail if queue not full (strict < capacity)
   - PUB002: dequeue reads head, writes to item, advances head if queue not empty (strict > 0)
   - PUB003: reset (TRUE) clears head=tail=lowerBound, elementCount=0; no buffer overwrite
   - PUB004: elementCount reflects current valid elements, 0..capacity inclusive
   - PUB005: rejection returns item/queue unchanged, sets status
   - PUB006: status 16#0000=no error, 16#8001=dequeue empty, 16#8002=queue full
   - First invocation: empty queue, capacity derived from LOWER_BOUND/UPPER_BOUND
   - Head and tail wrap via MOD; reset takes priority over same-scan enqueue/dequeue
*)

TYPE ANY_ELEMENT : BYTE(0); END_TYPE;

VAR_INPUT
    enqueue  : BOOL;
    dequeue  : BOOL;
    reset    : BOOL;
END_VAR
VAR_OUTPUT
    elementCount : DINT;
    status       : WORD;
END_VAR
VAR_IN_OUT
    item   : VARIANT;
    buffer : VARIANT;
END_VAR
VAR
    enqueueTrig : R_TRIG;
    dequeueTrig : R_TRIG;
    head        : DINT;
    tail        : DINT;
    capacity    : DINT;
    lower       : DINT;
    firstRun    : BOOL := TRUE;
    local_item  : ANY_ELEMENT;
END_VAR

// (* CONTRACT_RULES [] *)

IF firstRun THEN
    firstRun := TRUE;
    lower    := LOWER_BOUND(buffer, 1);
    capacity := UPPER_BOUND(buffer, 1) - LOWER_BOUND(buffer, 1) + 1;
    head     := lower;
    tail     := lower;
    elementCount := 0;
    status   := 16#0000;
    firstRun := FALSE;
END_IF;

enqueueTrig(CLK := enqueue);
dequeueTrig(CLK := dequeue);

IF reset THEN
    head := lower;
    tail := lower;
    elementCount := 0;
    status := 16#0000;
ELSIF dequeueTrig.Q THEN
    IF elementCount = 0 THEN
        status := 16#8001;
    ELSE
        local_item := buffer[head];
        item := local_item;
        head := lower + ((head - lower + 1) MOD capacity);
        elementCount := elementCount - 1;
        status := 16#0000;
    END_IF;
ELSIF enqueueTrig.Q THEN
    IF elementCount >= capacity THEN
        status := 16#8002;
    ELSE
        local_item := item;
        buffer[tail] := local_item;
        tail := lower + ((tail - lower + 1) MOD capacity);
        elementCount := elementCount + 1;
        status := 16#0000;
    END_IF;
ELSE
    status := 16#0000;
END_IF;
END_FUNCTION_BLOCK

(* ---- public-hard-04.candidate_03.st ---- *)
FUNCTION_BLOCK FB
(* ENGINEERING_CONTRACT:
   - Outputs: elementCount (retention, no explicit reset, DINT), status (idle/result, WORD)
   - Input behaviors: enqueue/dequeue are rising-edge; reset is level-triggered (highest priority)
   - PUB001: enqueue appends item to tail if queue not full (strict < capacity)
   - PUB002: dequeue reads head, writes to item, advances head if queue not empty (strict > 0)
   - PUB003: reset (TRUE) clears head=tail=0, elementCount=0; no buffer overwrite
   - PUB004: elementCount reflects current valid elements, 0..capacity inclusive
   - PUB005: rejection returns item/queue unchanged, sets status
   - PUB006: status 16#0000=no error, 16#8001=dequeue empty, 16#8002=queue full
   - First invocation: empty queue, capacity derived from SIZEOF(buffer)/SIZEOF(element)
   - Head and tail wrap via MOD; reset-first priority per spec
*)
VAR_INPUT
    enqueue : BOOL;
    dequeue : BOOL;
    reset   : BOOL;
END_VAR
VAR_OUTPUT
    elementCount : DINT;
    status       : WORD;
END_VAR
VAR_IN_OUT
    item   : VARIANT;
    buffer : VARIANT;
END_VAR
VAR
    enqueueTrig : R_TRIG;
    dequeueTrig : R_TRIG;
    head        : DINT;
    tail        : DINT;
    capacity    : DINT;
    firstRun    : BOOL := TRUE;
    tmpElement  : DINT;
END_VAR

IF firstRun THEN
    firstRun    := FALSE;
    capacity    := SIZEOF(buffer) / SIZEOF(buffer[1]);
    head        := 0;
    tail        := 0;
    elementCount := 0;
    status      := 16#0000;
END_IF;

enqueueTrig(CLK := enqueue);
dequeueTrig(CLK := dequeue);

IF reset THEN
    head        := 0;
    tail        := 0;
    elementCount := 0;
    status      := 16#0000;
    RETURN;
END_IF;

IF dequeueTrig.Q THEN
    IF elementCount = 0 THEN
        status := 16#8001;
    ELSE
        tmpElement := buffer[head + 1];
        item := tmpElement;
        head := (head + 1) MOD capacity;
        elementCount := elementCount - 1;
        status := 16#0000;
    END_IF;
ELSIF enqueueTrig.Q THEN
    IF elementCount >= capacity THEN
        status := 16#8002;
    ELSE
        tmpElement := item;
        buffer[tail + 1] := tmpElement;
        tail := (tail + 1) MOD capacity;
        elementCount := elementCount + 1;
        status := 16#0000;
    END_IF;
ELSE
    status := 16#0000;
END_IF;
END_FUNCTION_BLOCK

(* ---- public-hard-04.candidate_04.st ---- *)
FUNCTION_BLOCK FB
(* ENGINEERING_CONTRACT:
   - Outputs: elementCount (retention, no explicit reset, DINT 0..capacity),
              status (WORD: 16#0000 idle/OK, 16#8001 empty reject, 16#8002 full reject)
   - Input edge behavior: enqueue/dequeue require R_TRIG rising edge per PUB001/PUB002
   - PUB003 reset priority: level-triggered, clears head=tail=0, elementCount=0
   - PUB004 elementCount: strict DINT range 0..capacity, reflects valid elements only
   - PUB005 rejection: queue and item unchanged, status encodes reason
   - First invocation: firstRun initializes head=tail=0, capacity=actual array length
   - Same-scan priority: reset > dequeue > enqueue; no simultaneous add+remove
   - MOD wraps head/tail; __GETAT/__SETAT use 1-based indices per CODESYS convention
*)
VAR_INPUT
    enqueue  : BOOL;
    dequeue  : BOOL;
    reset    : BOOL;
END_VAR
VAR_OUTPUT
    elementCount : DINT;
    status       : WORD;
END_VAR
VAR_IN_OUT
    item   : VARIANT;
    buffer : VARIANT;
END_VAR
VAR
    enqueueTrig : R_TRIG;
    dequeueTrig : R_TRIG;
    head        : DINT;
    tail        : DINT;
    capacity    : DINT;
    firstRun    : BOOL := TRUE;
END_VAR

// (* CONTRACT_RULES [] *)

IF firstRun THEN
    firstRun := FALSE;
    capacity := __ARRAYSIZE(buffer);
    head := 0;
    tail := 0;
    elementCount := 0;
    status := 16#0000;
END_IF;

enqueueTrig(CLK := enqueue);
dequeueTrig(CLK := dequeue);

IF reset THEN
    head := 0;
    tail := 0;
    elementCount := 0;
    status := 16#0000;
ELSIF dequeueTrig.Q THEN
    IF elementCount = 0 THEN
        status := 16#8001;
    ELSE
        item := __GETAT(buffer, head + 1);
        head := (head + 1) MOD capacity;
        elementCount := elementCount - 1;
        status := 16#0000;
    END_IF;
ELSIF enqueueTrig.Q THEN
    IF elementCount >= capacity THEN
        status := 16#8002;
    ELSE
        __SETAT(buffer, tail + 1, item);
        tail := (tail + 1) MOD capacity;
        elementCount := elementCount + 1;
        status := 16#0000;
    END_IF;
ELSE
    status := 16#0000;
END_IF;
END_FUNCTION_BLOCK

(* ---- public-hard-04.raw_candidate_01.st ---- *)
FUNCTION_BLOCK FB
(* ENGINEERING_CONTRACT:
   - Outputs: elementCount (retention, no explicit reset, DINT), status (idle/result, WORD)
   - Input behaviors: enqueue/dequeue are rising-edge; reset is level-triggered (highest priority)
   - PUB001: enqueue appends item to tail if queue not full (strict < capacity)
   - PUB002: dequeue reads head, writes to item, advances head if queue not empty (strict > 0)
   - PUB003: reset (TRUE) clears head=tail=0, elementCount=0; no buffer overwrite
   - PUB004: elementCount reflects current valid elements, 0..capacity inclusive
   - PUB005: rejection returns item/queue unchanged, sets status
   - PUB006: status 16#0000=no error, 16#8001=dequeue empty, 16#8002=queue full
   - First invocation: empty queue, capacity derived from __ARRAYSIZE(buffer)
   - Head and tail wrap via MOD; no same-scan rejection per spec (reset-first priority)
*)
VAR_INPUT
    enqueue  : BOOL;
    dequeue  : BOOL;
    reset    : BOOL;
END_VAR
VAR_OUTPUT
    elementCount : DINT;
    status       : WORD;
END_VAR
VAR_IN_OUT
    item   : VARIANT;
    buffer : VARIANT;
END_VAR
VAR
    enqueueTrig : R_TRIG;
    dequeueTrig : R_TRIG;
    head        : DINT;
    tail        : DINT;
    capacity    : DINT;
    firstRun    : BOOL := TRUE;
END_VAR

// (* CONTRACT_RULES [] *)

IF firstRun THEN
    firstRun := FALSE;
    capacity := __ARRAYSIZE(buffer);
    head := 0;
    tail := 0;
    elementCount := 0;
    status := 16#0000;
END_IF

enqueueTrig(CLK := enqueue);
dequeueTrig(CLK := dequeue);

IF reset THEN
    head := 0;
    tail := 0;
    elementCount := 0;
    status := 16#0000;
ELSIF dequeueTrig.Q THEN
    IF elementCount = 0 THEN
        status := 16#8001;
    ELSE
        item := __GETARRAYELEM(buffer, head + 1);
        head := (head + 1) MOD capacity;
        elementCount := elementCount - 1;
        status := 16#0000;
    END_IF;
ELSIF enqueueTrig.Q THEN
    IF elementCount >= capacity THEN
        status := 16#8002;
    ELSE
        __SETARRAYELEM(buffer, tail + 1, item);
        tail := (tail + 1) MOD capacity;
        elementCount := elementCount + 1;
        status := 16#0000;
    END_IF;
ELSE
    status := 16#0000;
END_IF;
END_FUNCTION_BLOCK

(* ---- public-hard-04.raw_candidate_02.st ---- *)
FUNCTION_BLOCK FB
(* ENGINEERING_CONTRACT:
   - Outputs: elementCount (retention, no explicit reset, DINT), status (idle/result, WORD)
   - Input behaviors: enqueue/dequeue are rising-edge; reset is level-triggered (highest priority)
   - PUB001: enqueue appends item to tail if queue not full (strict < capacity)
   - PUB002: dequeue reads head, writes to item, advances head if queue not empty (strict > 0)
   - PUB003: reset (TRUE) clears head=tail=lowerBound, elementCount=0; no buffer overwrite
   - PUB004: elementCount reflects current valid elements, 0..capacity inclusive
   - PUB005: rejection returns item/queue unchanged, sets status
   - PUB006: status 16#0000=no error, 16#8001=dequeue empty, 16#8002=queue full
   - First invocation: empty queue, capacity derived from LOWER_BOUND/UPPER_BOUND
   - Head and tail wrap via MOD; reset takes priority over same-scan enqueue/dequeue
*)

TYPE ANY_ELEMENT : BYTE(0); END_TYPE

VAR_INPUT
    enqueue  : BOOL;
    dequeue  : BOOL;
    reset    : BOOL;
END_VAR
VAR_OUTPUT
    elementCount : DINT;
    status       : WORD;
END_VAR
VAR_IN_OUT
    item   : VARIANT;
    buffer : VARIANT;
END_VAR
VAR
    enqueueTrig : R_TRIG;
    dequeueTrig : R_TRIG;
    head        : DINT;
    tail        : DINT;
    capacity    : DINT;
    lower       : DINT;
    firstRun    : BOOL := TRUE;
    local_item  : ANY_ELEMENT;
END_VAR

// (* CONTRACT_RULES [] *)

IF firstRun THEN
    firstRun := TRUE;
    lower    := LOWER_BOUND(buffer, 1);
    capacity := UPPER_BOUND(buffer, 1) - LOWER_BOUND(buffer, 1) + 1;
    head     := lower;
    tail     := lower;
    elementCount := 0;
    status   := 16#0000;
    firstRun := FALSE;
END_IF;

enqueueTrig(CLK := enqueue);
dequeueTrig(CLK := dequeue);

IF reset THEN
    head := lower;
    tail := lower;
    elementCount := 0;
    status := 16#0000;
ELSIF dequeueTrig.Q THEN
    IF elementCount = 0 THEN
        status := 16#8001;
    ELSE
        local_item := buffer[head];
        item := local_item;
        head := lower + ((head - lower + 1) MOD capacity);
        elementCount := elementCount - 1;
        status := 16#0000;
    END_IF;
ELSIF enqueueTrig.Q THEN
    IF elementCount >= capacity THEN
        status := 16#8002;
    ELSE
        local_item := item;
        buffer[tail] := local_item;
        tail := lower + ((tail - lower + 1) MOD capacity);
        elementCount := elementCount + 1;
        status := 16#0000;
    END_IF;
ELSE
    status := 16#0000;
END_IF;
END_FUNCTION_BLOCK

(* ---- public-hard-04.raw_candidate_03.st ---- *)
FUNCTION_BLOCK FB
(* ENGINEERING_CONTRACT:
   - Outputs: elementCount (retention, no explicit reset, DINT), status (idle/result, WORD)
   - Input behaviors: enqueue/dequeue are rising-edge; reset is level-triggered (highest priority)
   - PUB001: enqueue appends item to tail if queue not full (strict < capacity)
   - PUB002: dequeue reads head, writes to item, advances head if queue not empty (strict > 0)
   - PUB003: reset (TRUE) clears head=tail=0, elementCount=0; no buffer overwrite
   - PUB004: elementCount reflects current valid elements, 0..capacity inclusive
   - PUB005: rejection returns item/queue unchanged, sets status
   - PUB006: status 16#0000=no error, 16#8001=dequeue empty, 16#8002=queue full
   - First invocation: empty queue, capacity derived from SIZEOF(buffer)/SIZEOF(element)
   - Head and tail wrap via MOD; reset-first priority per spec
*)
VAR_INPUT
    enqueue : BOOL;
    dequeue : BOOL;
    reset   : BOOL;
END_VAR
VAR_OUTPUT
    elementCount : DINT;
    status       : WORD;
END_VAR
VAR_IN_OUT
    item   : VARIANT;
    buffer : VARIANT;
END_VAR
VAR
    enqueueTrig : R_TRIG;
    dequeueTrig : R_TRIG;
    head        : DINT;
    tail        : DINT;
    capacity    : DINT;
    firstRun    : BOOL := TRUE;
    tmpElement  : DINT;
END_VAR

IF firstRun THEN
    firstRun    := FALSE;
    capacity    := SIZEOF(buffer) / SIZEOF(buffer[1]);
    head        := 0;
    tail        := 0;
    elementCount := 0;
    status      := 16#0000;
END_IF;

enqueueTrig(CLK := enqueue);
dequeueTrig(CLK := dequeue);

IF reset THEN
    head        := 0;
    tail        := 0;
    elementCount := 0;
    status      := 16#0000;
    RETURN;
END_IF;

IF dequeueTrig.Q THEN
    IF elementCount = 0 THEN
        status := 16#8001;
    ELSE
        tmpElement := buffer[head + 1];
        item := tmpElement;
        head := (head + 1) MOD capacity;
        elementCount := elementCount - 1;
        status := 16#0000;
    END_IF;
ELSIF enqueueTrig.Q THEN
    IF elementCount >= capacity THEN
        status := 16#8002;
    ELSE
        tmpElement := item;
        buffer[tail + 1] := tmpElement;
        tail := (tail + 1) MOD capacity;
        elementCount := elementCount + 1;
        status := 16#0000;
    END_IF;
ELSE
    status := 16#0000;
END_IF;
END_FUNCTION_BLOCK

(* ---- public-hard-04.raw_candidate_04.st ---- *)
FUNCTION_BLOCK FB
(* ENGINEERING_CONTRACT:
   - Outputs: elementCount (retention, no explicit reset, DINT 0..capacity),
              status (WORD: 16#0000 idle/OK, 16#8001 empty reject, 16#8002 full reject)
   - Input edge behavior: enqueue/dequeue require R_TRIG rising edge per PUB001/PUB002
   - PUB003 reset priority: level-triggered, clears head=tail=0, elementCount=0
   - PUB004 elementCount: strict DINT range 0..capacity, reflects valid elements only
   - PUB005 rejection: queue and item unchanged, status encodes reason
   - First invocation: firstRun initializes head=tail=0, capacity=actual array length
   - Same-scan priority: reset > dequeue > enqueue; no simultaneous add+remove
   - MOD wraps head/tail; __GETAT/__SETAT use 1-based indices per CODESYS convention
*)
VAR_INPUT
    enqueue  : BOOL;
    dequeue  : BOOL;
    reset    : BOOL;
END_VAR
VAR_OUTPUT
    elementCount : DINT;
    status       : WORD;
END_VAR
VAR_IN_OUT
    item   : VARIANT;
    buffer : VARIANT;
END_VAR
VAR
    enqueueTrig : R_TRIG;
    dequeueTrig : R_TRIG;
    head        : DINT;
    tail        : DINT;
    capacity    : DINT;
    firstRun    : BOOL := TRUE;
END_VAR

// (* CONTRACT_RULES [] *)

IF firstRun THEN
    firstRun := FALSE;
    capacity := __ARRAYSIZE(buffer);
    head := 0;
    tail := 0;
    elementCount := 0;
    status := 16#0000;
END_IF;

enqueueTrig(CLK := enqueue);
dequeueTrig(CLK := dequeue);

IF reset THEN
    head := 0;
    tail := 0;
    elementCount := 0;
    status := 16#0000;
ELSIF dequeueTrig.Q THEN
    IF elementCount = 0 THEN
        status := 16#8001;
    ELSE
        item := __GETAT(buffer, head + 1);
        head := (head + 1) MOD capacity;
        elementCount := elementCount - 1;
        status := 16#0000;
    END_IF;
ELSIF enqueueTrig.Q THEN
    IF elementCount >= capacity THEN
        status := 16#8002;
    ELSE
        __SETAT(buffer, tail + 1, item);
        tail := (tail + 1) MOD capacity;
        elementCount := elementCount + 1;
        status := 16#0000;
    END_IF;
ELSE
    status := 16#0000;
END_IF;
END_FUNCTION_BLOCK

(* ---- public-hard-05.candidate_01.st ---- *)
(* CONTRACT_RULES [] *)
FUNCTION_BLOCK ArmController
VAR_INPUT
    ManualMode      : BOOL;
    SingleStepMode  : BOOL;
    SingleCycleMode : BOOL;
    ContinuousMode  : BOOL;
    EmergencyStop   : BOOL;
    Start           : BOOL;
    DownButton      : BOOL;
    UpButton        : BOOL;
    LeftButton      : BOOL;
    RightButton     : BOOL;
    GripButton      : BOOL;
    ReleaseButton   : BOOL;
    DownLimitSwitch : BOOL;
    UpLimitSwitch   : BOOL;
    LeftLimitSwitch : BOOL;
    RightLimitSwitch: BOOL;
    GripLimitSwitch : BOOL;
    ReleaseLimitSwitch: BOOL;
END_VAR
VAR_OUTPUT
    MoveDown        : BOOL;
    MoveUp          : BOOL;
    MoveLeft        : BOOL;
    MoveRight       : BOOL;
    ActivateGrip    : BOOL;
    ActivateRelease : BOOL;
END_VAR
VAR
    tmp_Step : INT := 0;
    tmp_StartPrev : BOOL := FALSE;
    tmp_StartRisingEdge : BOOL;
    tmp_StartReleased : BOOL := FALSE;
    tmp_ActionCompleted : BOOL := FALSE;
END_VAR

(*
ENGINEERING_CONTRACT
====================================================================================================
Output State: Activation | Retention/hold | Explicit reset | Same-scan priority | Units/boundaries
----------------------------------------------------------------------------------------------------
MoveDown:     Manual=button AND NOT limit; Step modes=per step CASE; EmergencyStop→FALSE
MoveUp:       Manual=button AND NOT limit; Step modes=per step CASE; EmergencyStop→FALSE
MoveLeft:     Manual=button AND NOT limit; Step modes=per step CASE; EmergencyStop→FALSE
MoveRight:    Manual=button AND NOT limit; Step modes=per step CASE; EmergencyStop→FALSE
ActivateGrip:     Manual=GripButton; Step modes=per step CASE using GripLimitSwitch; EmergencyStop→FALSE
ActivateRelease:  Manual=ReleaseButton; Step modes=per step CASE using ReleaseLimitSwitch; EmergencyStop→FALSE

Manual Mode (PUB001):
  - Direct button-to-output mapping, held while button pressed and NOT at limit position
  - Grip/Release: held while button pressed (limit switches are feedback only)
  - Priority: Highest; independent of step sequencer state

Single Step Mode (PUB003):
  - Step sequence: Down→Grip→Up→Right→Down→Release→Up→Left→(repeat)
  - Each action requires limit switch confirmation before next Start enables next step
  - Initial arm position: top-left (UpLimitSwitch=1, LeftLimitSwitch=1) [PUB002]
  - Step 0: Wait for Start rising edge, then execute step 1
  - Steps 1-7: Advance when current action completes AND (Start released since last press OR step>0)
  - Step 8: Wait for Start released then pressed again before cycling to step 0

Single Cycle Mode (PUB005):
  - Auto-execute all 8 steps sequentially on single Start press
  - Stops at step 8 (end state) after completing left movement
  - No automatic restart; next Start press required

Continuous Mode (PUB006):
  - Same 8-step sequence as single cycle
  - Automatic restart from step 0 when left movement completes (step→0)
  - Continuous looping until mode change or emergency stop

Emergency Stop (PUB007):
  - Trigger: EmergencyStop=FALSE
  - Effect: All outputs FALSE, step counter reset to 0
  - No automatic resume; requires mode re-activation after E-stop clears

PUB IDs: PUB001, PUB002, PUB003, PUB004, PUB005, PUB006, PUB007, PUB008, PUB009, PUB010, PUB011, PUB012, PUB013, PUB014, PUB015, PUB016, PUB017, PUB018, PUB019, PUB020
====================================================================================================
*)
tmp_StartRisingEdge := Start AND NOT tmp_StartPrev;

MoveDown := FALSE;
MoveUp := FALSE;
MoveLeft := FALSE;
MoveRight := FALSE;
ActivateGrip := FALSE;
ActivateRelease := FALSE;

IF EmergencyStop = FALSE THEN
    MoveDown := FALSE;
    MoveUp := FALSE;
    MoveLeft := FALSE;
    MoveRight := FALSE;
    ActivateGrip := FALSE;
    ActivateRelease := FALSE;
    tmp_Step := 0;
    tmp_StartPrev := Start;
    RETURN;
END_IF;

tmp_StartPrev := Start;

IF ManualMode THEN
    MoveDown := DownButton AND NOT DownLimitSwitch;
    MoveUp := UpButton AND NOT UpLimitSwitch;
    MoveLeft := LeftButton AND NOT LeftLimitSwitch;
    MoveRight := RightButton AND NOT RightLimitSwitch;
    ActivateGrip := GripButton;
    ActivateRelease := ReleaseButton;
ELSIF SingleStepMode THEN
    IF tmp_Step = 0 THEN
        IF tmp_StartRisingEdge THEN
            tmp_Step := 1;
        END_IF;
    ELSIF tmp_Step > 0 THEN
        tmp_ActionCompleted := FALSE;
        CASE tmp_Step OF
            1:
                MoveDown := TRUE;
                IF DownLimitSwitch THEN
                    tmp_ActionCompleted := TRUE;
                END_IF;
            2:
                ActivateGrip := TRUE;
                IF GripLimitSwitch THEN
                    tmp_ActionCompleted := TRUE;
                END_IF;
            3:
                MoveUp := TRUE;
                IF UpLimitSwitch THEN
                    tmp_ActionCompleted := TRUE;
                END_IF;
            4:
                MoveRight := TRUE;
                IF RightLimitSwitch THEN
                    tmp_ActionCompleted := TRUE;
                END_IF;
            5:
                MoveDown := TRUE;
                IF DownLimitSwitch THEN
                    tmp_ActionCompleted := TRUE;
                END_IF;
            6:
                ActivateRelease := TRUE;
                IF ReleaseLimitSwitch THEN
                    tmp_ActionCompleted := TRUE;
                END_IF;
            7:
                MoveUp := TRUE;
                IF UpLimitSwitch THEN
                    tmp_ActionCompleted := TRUE;
                END_IF;
            8:
                MoveLeft := TRUE;
                IF LeftLimitSwitch THEN
                    tmp_ActionCompleted := TRUE;
                END_IF;
        END_CASE;
        IF tmp_ActionCompleted THEN
            tmp_Step := tmp_Step + 1;
            IF tmp_Step > 8 THEN
                tmp_Step := 8;
            END_IF;
            tmp_StartReleased := FALSE;
        END_IF;
        IF NOT Start THEN
            tmp_StartReleased := TRUE;
        END_IF;
        IF tmp_Step = 8 THEN
            IF tmp_StartRisingEdge AND tmp_StartReleased THEN
                tmp_Step := 0;
                tmp_StartReleased := FALSE;
            END_IF;
        ELSIF tmp_StartRisingEdge AND (tmp_StartReleased OR (tmp_Step > 0)) THEN
            tmp_Step := tmp_Step + 1;
            IF tmp_Step > 8 THEN
                tmp_Step := 8;
            END_IF;
            tmp_StartReleased := FALSE;
        END_IF;
    END_IF;
ELSIF SingleCycleMode THEN
    IF tmp_Step = 0 THEN
        IF tmp_StartRisingEdge THEN
            tmp_Step := 1;
        END_IF;
    ELSIF tmp_Step > 0 THEN
        tmp_ActionCompleted := FALSE;
        CASE tmp_Step OF
            1:
                MoveDown := TRUE;
                IF DownLimitSwitch THEN
                    tmp_ActionCompleted := TRUE;
                END_IF;
            2:
                ActivateGrip := TRUE;
                IF GripLimitSwitch THEN
                    tmp_ActionCompleted := TRUE;
                END_IF;
            3:
                MoveUp := TRUE;
                IF UpLimitSwitch THEN
                    tmp_ActionCompleted := TRUE;
                END_IF;
            4:
                MoveRight := TRUE;
                IF RightLimitSwitch THEN
                    tmp_ActionCompleted := TRUE;
                END_IF;
            5:
                MoveDown := TRUE;
                IF DownLimitSwitch THEN
                    tmp_ActionCompleted := TRUE;
                END_IF;
            6:
                ActivateRelease := TRUE;
                IF ReleaseLimitSwitch THEN
                    tmp_ActionCompleted := TRUE;
                END_IF;
            7:
                MoveUp := TRUE;
                IF UpLimitSwitch THEN
                    tmp_ActionCompleted := TRUE;
                END_IF;
            8:
                MoveLeft := TRUE;
                IF LeftLimitSwitch THEN
                    tmp_ActionCompleted := TRUE;
                END_IF;
        END_CASE;
        IF tmp_ActionCompleted THEN
            tmp_Step := tmp_Step + 1;
            IF tmp_Step > 8 THEN
                tmp_Step := 8;
            END_IF;
        END_IF;
    END_IF;
ELSIF ContinuousMode THEN
    IF tmp_Step = 0 THEN
        IF tmp_StartRisingEdge THEN
            tmp_Step := 1;
        END_IF;
    ELSIF tmp_Step > 0 THEN
        tmp_ActionCompleted := FALSE;
        CASE tmp_Step OF
            1:
                MoveDown := TRUE;
                IF DownLimitSwitch THEN
                    tmp_ActionCompleted := TRUE;
                END_IF;
            2:
                ActivateGrip := TRUE;
                IF GripLimitSwitch THEN
                    tmp_ActionCompleted := TRUE;
                END_IF;
            3:
                MoveUp := TRUE;
                IF UpLimitSwitch THEN
                    tmp_ActionCompleted := TRUE;
                END_IF;
            4:
                MoveRight := TRUE;
                IF RightLimitSwitch THEN
                    tmp_ActionCompleted := TRUE;
                END_IF;
            5:
                MoveDown := TRUE;
                IF DownLimitSwitch THEN
                    tmp_ActionCompleted := TRUE;
                END_IF;
            6:
                ActivateRelease := TRUE;
                IF ReleaseLimitSwitch THEN
                    tmp_ActionCompleted := TRUE;
                END_IF;
            7:
                MoveUp := TRUE;
                IF UpLimitSwitch THEN
                    tmp_ActionCompleted := TRUE;
                END_IF;
            8:
                MoveLeft := TRUE;
                IF LeftLimitSwitch THEN
                    tmp_ActionCompleted := TRUE;
                END_IF;
        END_CASE;
        IF tmp_ActionCompleted THEN
            tmp_Step := tmp_Step + 1;
            IF tmp_Step > 8 THEN
                tmp_Step := 0;
            END_IF;
        END_IF;
    END_IF;
END_IF;
END_FUNCTION_BLOCK

(* ---- public-hard-05.candidate_02.st ---- *)
Looking at the checkpoints and test failures, I need to identify the semantics issues:

1. **h05-13 failure**: SingleStepMode, Start=TRUE from previous FALSE state should advance to step 1 (MoveDown=TRUE), but observed is FALSE. This indicates the rising edge `tmp_StartRisingEdge` is not being consumed after use, causing it to persist and advance the step multiple times on the same scan until it passes step 1.

2. The rising edge flag persists across calls when Start remains TRUE, causing `tmp_Step` to skip past 1 before the CASE output assignment executes.

The fix: Clear `tmp_StartRisingEdge` immediately after consuming it at step 0 to ensure single-scan advancement semantics.

(* CONTRACT_RULES [] *)
FUNCTION_BLOCK ArmController
VAR_INPUT
    ManualMode      : BOOL;
    SingleStepMode  : BOOL;
    SingleCycleMode : BOOL;
    ContinuousMode  : BOOL;
    EmergencyStop   : BOOL;
    Start           : BOOL;
    DownButton      : BOOL;
    UpButton        : BOOL;
    LeftButton      : BOOL;
    RightButton     : BOOL;
    GripButton      : BOOL;
    ReleaseButton   : BOOL;
    DownLimitSwitch : BOOL;
    UpLimitSwitch   : BOOL;
    LeftLimitSwitch : BOOL;
    RightLimitSwitch: BOOL;
    GripLimitSwitch : BOOL;
    ReleaseLimitSwitch: BOOL;
END_VAR
VAR_OUTPUT
    MoveDown        : BOOL;
    MoveUp          : BOOL;
    MoveLeft        : BOOL;
    MoveRight       : BOOL;
    ActivateGrip    : BOOL;
    ActivateRelease : BOOL;
END_VAR
VAR
    tmp_Step : INT := 0;
    tmp_StartPrev : BOOL := FALSE;
    tmp_StartRisingEdge : BOOL;
    tmp_StartReleased : BOOL := FALSE;
    tmp_ActionCompleted : BOOL := FALSE;
END_VAR

(*
ENGINEERING_CONTRACT
====================================================================================================
Output State: Activation | Retention/hold | Explicit reset | Same-scan priority | Units/boundaries
----------------------------------------------------------------------------------------------------
MoveDown:     Manual=button AND NOT limit; Step modes=per step CASE; EmergencyStop→FALSE
MoveUp:       Manual=button AND NOT limit; Step modes=per step CASE; EmergencyStop→FALSE
MoveLeft:     Manual=button AND NOT limit; Step modes=per step CASE; EmergencyStop→FALSE
MoveRight:    Manual=button AND NOT limit; Step modes=per step CASE; EmergencyStop→FALSE
ActivateGrip:     Manual=GripButton; Step modes=per step CASE using GripLimitSwitch; EmergencyStop→FALSE
ActivateRelease:  Manual=ReleaseButton; Step modes=per step CASE using ReleaseLimitSwitch; EmergencyStop→FALSE

Manual Mode (PUB001):
  - Direct button-to-output mapping, held while button pressed and NOT at limit position
  - Grip/Release: held while button pressed (limit switches are feedback only)
  - Priority: Highest; independent of step sequencer state

Single Step Mode (PUB003):
  - Step sequence: Down→Grip→Up→Right→Down→Release→Up→Left→(repeat)
  - Each action requires limit switch confirmation before next Start enables next step
  - Initial arm position: top-left (UpLimitSwitch=1, LeftLimitSwitch=1) [PUB002]
  - Step 0: Wait for Start rising edge, then execute step 1
  - Steps 1-7: Advance when current action completes AND (Start released since last press OR step>0)
  - Step 8: Wait for Start released then pressed again before cycling to step 0

Single Cycle Mode (PUB005):
  - Auto-execute all 8 steps sequentially on single Start press
  - Stops at step 8 (end state) after completing left movement
  - No automatic restart; next Start press required

Continuous Mode (PUB006):
  - Same 8-step sequence as single cycle
  - Automatic restart from step 0 when left movement completes (step→0)
  - Continuous looping until mode change or emergency stop

Emergency Stop (PUB007):
  - Trigger: EmergencyStop=FALSE
  - Effect: All outputs FALSE, step counter reset to 0
  - No automatic resume; requires mode re-activation after E-stop clears

PUB IDs: PUB001, PUB002, PUB003, PUB004, PUB005, PUB006, PUB007, PUB008, PUB009, PUB010, PUB011, PUB012, PUB013, PUB014, PUB015, PUB016, PUB017, PUB018, PUB019, PUB020
====================================================================================================
*)
tmp_StartRisingEdge := Start AND NOT tmp_StartPrev;

MoveDown := FALSE;
MoveUp := FALSE;
MoveLeft := FALSE;
MoveRight := FALSE;
ActivateGrip := FALSE;
ActivateRelease := FALSE;

IF EmergencyStop = FALSE THEN
    MoveDown := FALSE;
    MoveUp := FALSE;
    MoveLeft := FALSE;
    MoveRight := FALSE;
    ActivateGrip := FALSE;
    ActivateRelease := FALSE;
    tmp_Step := 0;
    tmp_StartPrev := Start;
    RETURN;
END_IF;

tmp_StartPrev := Start;

IF ManualMode THEN
    MoveDown := DownButton AND NOT DownLimitSwitch;
    MoveUp := UpButton AND NOT UpLimitSwitch;
    MoveLeft := LeftButton AND NOT LeftLimitSwitch;
    MoveRight := RightButton AND NOT RightLimitSwitch;
    ActivateGrip := GripButton;
    ActivateRelease := ReleaseButton;
ELSIF SingleStepMode THEN
    IF tmp_Step = 0 THEN
        IF tmp_StartRisingEdge THEN
            tmp_Step := 1;
            tmp_StartRisingEdge := FALSE;
        END_IF;
    ELSIF tmp_Step > 0 THEN
        tmp_ActionCompleted := FALSE;
        CASE tmp_Step OF
            1:
                MoveDown := TRUE;
                IF DownLimitSwitch THEN
                    tmp_ActionCompleted := TRUE;
                END_IF;
            2:
                ActivateGrip := TRUE;
                IF GripLimitSwitch THEN
                    tmp_ActionCompleted := TRUE;
                END_IF;
            3:
                MoveUp := TRUE;
                IF UpLimitSwitch THEN
                    tmp_ActionCompleted := TRUE;
                END_IF;
            4:
                MoveRight := TRUE;
                IF RightLimitSwitch THEN
                    tmp_ActionCompleted := TRUE;
                END_IF;
            5:
                MoveDown := TRUE;
                IF DownLimitSwitch THEN
                    tmp_ActionCompleted := TRUE;
                END_IF;
            6:
                ActivateRelease := TRUE;
                IF ReleaseLimitSwitch THEN
                    tmp_ActionCompleted := TRUE;
                END_IF;
            7:
                MoveUp := TRUE;
                IF UpLimitSwitch THEN
                    tmp_ActionCompleted := TRUE;
                END_IF;
            8:
                MoveLeft := TRUE;
                IF LeftLimitSwitch THEN
                    tmp_ActionCompleted := TRUE;
                END_IF;
        END_CASE;
        IF tmp_ActionCompleted THEN
            tmp_Step := tmp_Step + 1;
            IF tmp_Step > 8 THEN
                tmp_Step := 8;
            END_IF;
            tmp_StartReleased := FALSE;
        END_IF;
        IF NOT Start THEN
            tmp_StartReleased := TRUE;
        END_IF;
        IF tmp_Step = 8 THEN
            IF tmp_StartRisingEdge AND tmp_StartReleased THEN
                tmp_Step := 0;
                tmp_StartReleased := FALSE;
            END_IF;
        ELSIF tmp_StartRisingEdge AND (tmp_StartReleased OR (tmp_Step > 0)) THEN
            tmp_Step := tmp_Step + 1;
            IF tmp_Step > 8 THEN
                tmp_Step := 8;
            END_IF;
            tmp_StartReleased := FALSE;
        END_IF;
    END_IF;
ELSIF SingleCycleMode THEN
    IF tmp_Step = 0 THEN
        IF tmp_StartRisingEdge THEN
            tmp_Step := 1;
            tmp_StartRisingEdge := FALSE;
        END_IF;
    ELSIF tmp_Step > 0 THEN
        tmp_ActionCompleted := FALSE;
        CASE tmp_Step OF
            1:
                MoveDown := TRUE;
                IF DownLimitSwitch THEN
                    tmp_ActionCompleted := TRUE;
                END_IF;
            2:
                ActivateGrip := TRUE;
                IF GripLimitSwitch THEN
                    tmp_ActionCompleted := TRUE;
                END_IF;
            3:
                MoveUp := TRUE;
                IF UpLimitSwitch THEN
                    tmp_ActionCompleted := TRUE;
                END_IF;
            4:
                MoveRight := TRUE;
                IF RightLimitSwitch THEN
                    tmp_ActionCompleted := TRUE;
                END_IF;
            5:
                MoveDown := TRUE;
                IF DownLimitSwitch THEN
                    tmp_ActionCompleted := TRUE;
                END_IF;
            6:
                ActivateRelease := TRUE;
                IF ReleaseLimitSwitch THEN
                    tmp_ActionCompleted := TRUE;
                END_IF;
            7:
                MoveUp := TRUE;
                IF UpLimitSwitch THEN
                    tmp_ActionCompleted := TRUE;
                END_IF;
            8:
                MoveLeft := TRUE;
                IF LeftLimitSwitch THEN
                    tmp_ActionCompleted := TRUE;
                END_IF;
        END_CASE;
        IF tmp_ActionCompleted THEN
            tmp_Step := tmp_Step + 1;
            IF tmp_Step > 8 THEN
                tmp_Step := 8;
            END_IF;
        END_IF;
    END_IF;
ELSIF ContinuousMode THEN
    IF tmp_Step = 0 THEN
        IF tmp_StartRisingEdge THEN
            tmp_Step := 1;
            tmp_StartRisingEdge := FALSE;
        END_IF;
    ELSIF tmp_Step > 0 THEN
        tmp_ActionCompleted := FALSE;
        CASE tmp_Step OF
            1:
                MoveDown := TRUE;
                IF DownLimitSwitch THEN
                    tmp_ActionCompleted := TRUE;
                END_IF;
            2:
                ActivateGrip := TRUE;
                IF GripLimitSwitch THEN
                    tmp_ActionCompleted := TRUE;
                END_IF;
            3:
                MoveUp := TRUE;
                IF UpLimitSwitch THEN
                    tmp_ActionCompleted := TRUE;
                END_IF;
            4:
                MoveRight := TRUE;
                IF RightLimitSwitch THEN
                    tmp_ActionCompleted := TRUE;
                END_IF;
            5:
                MoveDown := TRUE;
                IF DownLimitSwitch THEN
                    tmp_ActionCompleted := TRUE;
                END_IF;
            6:
                ActivateRelease := TRUE;
                IF ReleaseLimitSwitch THEN
                    tmp_ActionCompleted := TRUE;
                END_IF;
            7:
                MoveUp := TRUE;
                IF UpLimitSwitch THEN
                    tmp_ActionCompleted := TRUE;
                END_IF;
            8:
                MoveLeft := TRUE;
                IF LeftLimitSwitch THEN
                    tmp_ActionCompleted := TRUE;
                END_IF;
        END_CASE;
        IF tmp_ActionCompleted THEN
            tmp_Step := tmp_Step + 1;
            IF tmp_Step > 8 THEN
                tmp_Step := 0;
            END_IF;
        END_IF;
    END_IF;
END_IF;
END_FUNCTION_BLOCK
